(* IEC 61131-3 sources: daoli-st-library/DL_Process (part 44) *)

(* ---- FB_DL_PalletizerLayerSeq.st ---- *)
//==============================================================================
// 功能块：FB_DL_PalletizerLayerSeq ｜ 中文名称：码垛层排布顺控
// 所属子库：DL_Process ｜ 版本：v1.0.1 ｜ 兼容：CODESYS V3.5+ / TwinCAT 3 / 汇川 InoProShop
// 功能描述：码垛机层排布顺控：层容量自算（正交与旋转两取向各算一遍，逐层按本层取向校验）→ 层内位置
//           序列 → 取放指令与夹手完成反馈握手（超时重试一次）→ 层满/垛满判定。
//           奇偶层旋转时偶数层整体旋转 90 度，层内落点由 FC_DL_Affine2Apply 施加旋转
//           矩阵得到（库内低层复用，禁止在本件重写点变换与矩阵乘）。旋转矩阵的元素以
//           VAR CONSTANT 标量常量声明（恒等 1/0、90 度 0/-1/+1），每拍装配成生效阵；
//           平移列恒为 0，运行时平移量（托盘长度）在阵外补偿——阵中不含运行时量，才配
//           得上常量语义（二维数组行主序字面量初始化在三平台可移植性差，故用标量常量
//           装配，避免方言差异）。本件只出位姿与指令，不做轨迹规划、不控夹手电磁阀
//           （执行器归设备层）。
// 开源溯源 (Origin)：道莅原创实现（参考 公开工程惯例 分类与参数域）
// 单位表：托盘与箱体尺寸[mm] / 层高[mm] / 坐标[mm] / 旋转角[度] / 层数与位置序号[个] /
//         取放超时[s] / 扫描间隔[ms] / 垛计数[垛]
// 错误码表：16#0005_0408 信息级（末层不满垛，留空位，不置 bError）/ 16#0005_0409 信息级
//           （取放超时首次重试，不置 bError）/ 16#0005_034E 故障级（层容量不足或箱体/
//           托盘尺寸规格不匹配，含尺寸非有限——非有限尺寸即规格不可信，映射见本行）/
//           16#0005_034F 故障级（取放超时重试耗尽，垛型中断，置 bError + 撤指令）/
//           16#0005_0350 故障级兜底（状态机落 ELSE 非法状态，置 bError）。034E 非有限
//           映射的反证句：尺寸非有限与容量不足在现有输出组合下不可观测出差异（均为
//           bError + bPlaceCmd 撤 + bValid 撤 + eState 进 eFault），§3 未给本件独立非有限
//           槽，故显式复用不越段。
// 状态机：E_DL_PalletLayerState（eIdle=0 待机 / eWaitCase=10 等来料 / ePlace=20 出取放
//           指令 / eWaitGrip=30 等夹手反馈 / eLayerEnd=40 层边界 / ePalletEnd=50 垛边界 /
//           eFault=99 故障兜底），CASE 含 ELSE 兜底，ELSE 置 0350 且撤指令、许可撤。
// 边界行为：① 层容量自算：正交取向 floor(托盘长/箱长) x floor(托盘宽/箱宽)、旋转取向
//           floor(托盘长/箱宽) x floor(托盘宽/箱长)，两取向各自校验——nCasePerLayer 超
//           正交容量 → 故障 034E；启用奇偶层旋转时还须不超旋转容量，否则同样 034E
//           （取大者会让旋转层"蒙混过关"，故逐取向验，绝不硬塞）；② 取放超时先重试
//           一次（信息 0409），二次超时 → 故障 034F 并中断垛型；③ 层高累计 Z =
//           (层号 − 1) x 层高，LREAL 承载防溢出；④ 末层不满 → 信息 0408；⑤ bStop 只在
//           层边界与等来料相生效（不在抓取中停，安全侧）；⑥ 失能/停止 → 撤指令 +
//           bValid := FALSE（R72）；⑦ 旋转落点必须走 FC_DL_Affine2Apply（常量纯旋转阵，
//           平移在阵外补偿），点变换件返回不可用 → 034E 并撤指令。
// 修订历史：v1.0.0 2026-11-17 首版（R25 派单 · §4.16，依赖 §4.2 件 FC_DL_Affine2Apply 语义）
//           v1.0.1 2026-11-17 终审修正两处（对外引脚契约零变更）：①旋转层阵外平移量由 fPalletLengthMm
//           改为 (nRowsEff − 1) x fCaseWidthMm（原式整体多推一个箱宽，首行落点越出托盘边界）；
//           ②bPalletDone 取消本相同拍自撤，撤销点移交 eIdle 相（原实现同拍置位又撤位，脉冲永不外显）。
//           层容量口径经总监独立验算：1200x1000 托盘配 400x300 箱体 → 正交 3x3=9、旋转 4x2=8，
//           派单书 §4.16 验收向量①所写「容量 6」为派单算术笔误，本件实现（9）为准。
//==============================================================================
(*------------------------------------------------------------------------------
 * 枚举: E_DL_PalletLayerState（归属 DL_Process，与 FB_DL_PalletizerLayerSeq 同文件）
 *----------------------------------------------------------------------------*)
TYPE E_DL_PalletLayerState :
(
    eIdle      := 0,   // 待机：指令撤，等 bStart / Idle, command dropped, waiting for start
    eWaitCase  := 10,  // 等来料：本层下一格位已算好，等 bCaseReady / Waiting for the next case
    ePlace     := 20,  // 出指令：bPlaceCmd 置位，等夹手动作 / Command issued, gripper acting
    eWaitGrip  := 30,  // 等反馈：等 bGripDone 或超时 / Waiting for feedback or timeout
    eLayerEnd  := 40,  // 层边界：本层放满，允许在此停止 / Layer boundary, a safe stop point
    ePalletEnd := 50,  // 垛边界：整垛完成，垛计数 +1 / Pallet boundary, pallet counter increments
    eFault     := 99   // 故障兜底：规格不匹配/超时耗尽/非法状态 / Fault fallback
);
END_TYPE

(*==============================================================================
 * 功能块: FB_DL_PalletizerLayerSeq
 * 调用约定: 每个扫描周期无条件调用一次；uDeltaTimeMs 必须注入真实任务间隔。
 *============================================================================*)
FUNCTION_BLOCK FB_DL_PalletizerLayerSeq
VAR_INPUT
    nCasePerLayer    : INT;                        // 每层箱数 [个]，须 <= 层容量 / Cases per layer [pcs], must not exceed the capacity
    nLayersPerPallet : INT;                        // 每垛层数 [层]，合法域 1~20 / Layers per pallet [layers], domain 1..20
    fPalletLengthMm  : LREAL;                      // 托盘长度 [mm]，须 > 0 / Pallet length [mm], must be > 0
    fPalletWidthMm   : LREAL;                      // 托盘宽度 [mm]，须 > 0 / Pallet width [mm], must be > 0
    fCaseLengthMm    : LREAL;                      // 箱体长度 [mm]，须 > 0 / Case length [mm], must be > 0
    fCaseWidthMm     : LREAL;                      // 箱体宽度 [mm]，须 > 0 / Case width [mm], must be > 0
    fLayerHeightMm   : LREAL;                      // 层高 [mm]，须 > 0 / Layer height [mm], must be > 0
    bOddLayerRotate  : BOOL;                       // 奇偶层旋转使能（偶数层旋转 90 度）/ Odd/even layer rotation, even layers rotate 90 degrees
    bCaseReady       : BOOL;                       // 来料在位 / Case available at the pick point
    bGripDone        : BOOL;                       // 夹手完成反馈 / Gripper completion feedback
    tGripTimeout     : TIME := T#8S;               // 取放超时 [ms] / Pick-and-place timeout [ms]
    bStart           : BOOL;                       // 启动（取上升沿）/ Start, rising edge
    bStop            : BOOL;                       // 停止（只在层边界与等来料相生效）/ Stop, honoured only at layer boundaries and while waiting
    bReset           : BOOL;                       // 复位，上升沿回待机并清垛计数锁存位 / Reset, rising edge returns to idle
    uDeltaTimeMs     : UDINT;                      // 扫描间隔 [ms]，调用方注入，禁系统时间函数 / Scan interval [ms], caller-injected
END_VAR
VAR_OUTPUT
    nLayerIndex      : INT;                        // 当前层号 [层]，从 1 起 / Current layer index, 1-based
    nPosIndex        : INT;                        // 层内位置序号 [个]，从 1 起 / In-layer position index, 1-based
    fTargetXMm       : LREAL;                      // 目标位 X [mm] / Target X [mm]
    fTargetYMm       : LREAL;                      // 目标位 Y [mm] / Target Y [mm]
    fTargetZMm       : LREAL;                      // 目标位 Z [mm] / Target Z [mm]
    fTargetRotDeg    : LREAL;                      // 目标旋转角 [度]，0 或 90 / Target rotation [deg], 0 or 90
    bPlaceCmd        : BOOL;                       // 取放指令（层放满/故障/停止即撤）/ Pick-and-place command
    bLayerDone       : BOOL;                       // 本层已放满 / Layer completed
    bPalletDone      : BOOL;                       // 整垛完成 / Pallet completed
    nCaseCount       : INT;                        // 本垛已放件数 [件] / Cases placed on this pallet [pcs]
    uPalletCount     : UDINT;                      // 完成垛数 [垛]，饱和 / Completed pallets [pallets], saturating
    eErr             : UDINT;                      // 错误码，0 = 无错，码位 16#0005_0408 起信息级、16#0005_034E 起故障级（分带见错误码表） / Error code, 0 = no error, band info/fault per the code table
    bError           : BOOL;                       // 故障级标志，仅故障级错误置位 / Fault-class flag, set only on fault-level codes
    bValid           : BOOL;                       // 位姿输出可用标志，失能/故障闸显式 FALSE / Pose usable flag, explicit FALSE on disable/fault gates
    eState           : E_DL_PalletLayerState;      // 主状态机当前状态 / Current state of the main state machine
END_VAR
VAR
    fbReset          : R_TRIG;                     // 复位上升沿检测实例 / Reset rising edge detector
    fbStart          : R_TRIG;                     // 启动上升沿检测实例 / Start rising edge detector
    fbTonGrip        : TON;                        // 取放超时定时器实例 / Pick-and-place timeout timer
    afRotZero        : ARRAY[0..2, 0..2] OF LREAL; // 本拍生效旋转矩阵（恒等或 90 度）/ Effective rotation matrix of this scan
    nCapOrtho        : INT;                        // 正交取向层容量 [件] / Capacity with the orthogonal orientation [pcs]
    nCapRot          : INT;                        // 旋转取向层容量 [件] / Capacity with the rotated orientation [pcs]
    nCapEff          : INT;                        // 本层取向容量 [件] / Capacity of the current orientation [pcs]
    nColsEff         : INT;                        // 本层列数 [个] / Columns of this layer [pcs]
    nRowsEff         : INT;                        // 本层行数 [个] / Rows of this layer [pcs]
    nIdx0            : INT;                        // 层内零基位置序号 [—] / Zero-based in-layer index
    nCol             : INT;                        // 本格位列号（1 基）[列] / Column of this cell, 1-based
    nRow             : INT;                        // 本格位行号（1 基）[行] / Row of this cell, 1-based
    nRetryCnt        : INT;                        // 本格位超时重试次数 [次] / Timeout retry count of this cell
    nLoop            : INT;                        // 赋值循环索引 [—] / Assignment loop index
    fLocalXMm        : LREAL;                      // 箱体自身坐标系 X [mm] / X in the case-local frame [mm]
    fLocalYMm        : LREAL;                      // 箱体自身坐标系 Y [mm] / Y in the case-local frame [mm]
    fOutXMm          : LREAL;                      // 点变换结果 X [mm] / Transformed X [mm]
    fOutYMm          : LREAL;                      // 点变换结果 Y [mm] / Transformed Y [mm]
    uApplyErr        : UDINT;                      // 点变换件错误码暂存 / Point-transform error code staging
    bApplyFault      : BOOL;                       // 点变换件故障标志暂存 / Point-transform fault flag staging
    bApplyValid      : BOOL;                       // 点变换件可用标志暂存 / Point-transform usable flag staging
    bApplyOk         : BOOL;                       // 点变换件返回值暂存 / Point-transform return staging
    bLayerRotated    : BOOL;                       // 本层旋转标志 / This layer is rotated
    bSpaceWarn       : BOOL;                       // 末层不满提示标志 / Under-filled top layer hint
    bGripTimedOut    : BOOL;                       // 取放超时命中 / Pick-and-place timeout hit
    bRearm           : BOOL;                       // 定时器重装脉冲（本拍强制 IN 为 FALSE 一拍）/ Timer re-arm pulse, forces IN FALSE for one scan
    bNonFin          : BOOL;                       // 非有限判定中间标志 / Non-finite detection intermediate flag
    bFirstScan       : BOOL := TRUE;               // 上电首拍标志 / First-scan flag
END_VAR
VAR CONSTANT
    DL_PLS_CODE_INFO_1 : UDINT := 16#0005_0408;    // 信息级槽 1（末层不满垛留空位） / info slot 1
    DL_PLS_CODE_INFO_2 : UDINT := 16#0005_0409;    // 信息级槽 2（取放超时重试） / info slot 2
    DL_PLS_CODE_FLT_1  : UDINT := 16#0005_034E;    // 故障级槽 1（容量不足/规格不匹配） / fault slot 1
    DL_PLS_CODE_FLT_2  : UDINT := 16#0005_034F;    // 故障级槽 2（超时重试耗尽） / fault slot 2
    DL_PLS_CODE_FLT_3  : UDINT := 16#0005_0350;    // 故障级槽 3（非法状态兜底） / fault slot 3, illegal-state fallback
    DL_PLS_ROT90       : LREAL := 90.0;            // 旋转层目标角 [度] / Rotated layer angle [deg]
    DL_PLS_LAYER_MIN   : INT := 1;                 // 层数下限 [层] / Layer count floor
    DL_PLS_LAYER_MAX   : INT := 20;                // 层数上限 [层] / Layer count ceiling
    DL_PLS_CELL_MIN    : INT := 1;                 // 层容量下限 [件] / Layer capacity floor [pcs]
    DL_PLS_CNT_MAX     : UDINT := 16#FFFF_FFFE;    // 垛计数饱和值 [垛] / Pallet counter saturation
    DL_PLS_RETRY_MAX   : INT := 1;                 // 超时重试次数上限 [次] / Retry ceiling [times]
    DL_PLS_ZERO        : LREAL := 0.0;             // 零值常量，避免裸字面量 [—] / Zero constant, avoids a bare literal
    DL_PLS_ONE         : LREAL := 1.0;             // 单位常量，齐次项 [—] / Unity constant, homogeneous entry
    DL_PLS_TOL         : LREAL := 1.0E-6;          // 浮点比较容差 [—] / Float comparison tolerance
    DL_PLS_INF         : LREAL := 1.7976931348623157E308; // LREAL 幅值上限，Inf 判据 / LREAL magnitude ceiling
    // 纯旋转常量阵（行主序平铺展开）：恒等映射 / pure rotation constants, row-major flat
    DL_PLS_M_ID_X      : LREAL := 1.0;             // 恒等阵 (0,0) / identity (0,0)
    DL_PLS_M_ID_Y      : LREAL := 1.0;             // 恒等阵 (1,1) / identity (1,1)
    DL_PLS_M_R90_C     : LREAL := -1.0;            // 90 度阵 (0,1) = -1 / rot90 (0,1) = -1
    DL_PLS_M_R90_S     : LREAL := 1.0;             // 90 度阵 (1,0) = +1 / rot90 (1,0) = +1
END_VAR

(*------------------------------------------------------------------------------
 * 段 1｜无条件刷新区（红线 5）：复位/启动沿与超时定时器在任意分支之外周期调用；
 *       定时器 IN 取上拍状态（单拍滞后对 8 s 窗无影响），保证各分支计时链不断流
 *----------------------------------------------------------------------------*)
fbReset(CLK := bReset);                            // 复位沿检测无条件刷新 / reset edge refreshed unconditionally
fbStart(CLK := bStart);                            // 启动沿检测无条件刷新 / start edge refreshed unconditionally
fbTonGrip(IN := (eState = E_DL_PalletLayerState.eWaitGrip) AND (NOT bGripDone)
                AND (NOT bRearm),                  // 重装拍强制 IN 为 FALSE 使定时器复位 / the re-arm scan forces IN FALSE, resetting the timer
          PT := tGripTimeout);                     // 取放超时 [ms] / pick-and-place timeout
IF bRearm THEN
    bRearm := FALSE;                               // 重装脉冲单拍自清（下一拍起重新计时）/ re-arm pulse self-cleared, timing restarts next scan
END_IF

(*------------------------------------------------------------------------------
 * 段 2｜复位沿处理（改写置于沿后，防吞沿 R39）
 *----------------------------------------------------------------------------*)
IF fbReset.Q THEN
    eState := E_DL_PalletLayerState.eIdle;
    eErr   := 16#0000_0000;                        // 复位清码 / reset clears the code
    bError := FALSE;                               // 复位清故障 / reset clears the fault
    nLayerIndex := 0;                              // 层号清 / layer index cleared
    nPosIndex := 0;                                // 位置序号清 / position index cleared
    nCaseCount := 0;                               // 本垛件数清 / pallet case count cleared
    nRetryCnt := 0;                                // 重试计数清 / retry count cleared
    bPlaceCmd := FALSE;                            // 指令撤 / command dropped
    bFirstScan := TRUE;                            // 重新首拍化 / re-initialize first scan
END_IF

(*------------------------------------------------------------------------------
 * 段 3｜非有限输入闸（尺寸类，R79）：映射入 034E（规格不可信，见错误码表反证句）
 *----------------------------------------------------------------------------*)
bNonFin := (fPalletLengthMm <> fPalletLengthMm) OR (ABS(fPalletLengthMm) >= DL_PLS_INF)
        OR (fPalletWidthMm <> fPalletWidthMm) OR (ABS(fPalletWidthMm) >= DL_PLS_INF)
        OR (fCaseLengthMm <> fCaseLengthMm) OR (ABS(fCaseLengthMm) >= DL_PLS_INF)
        OR (fCaseWidthMm <> fCaseWidthMm) OR (ABS(fCaseWidthMm) >= DL_PLS_INF)
        OR (fLayerHeightMm <> fLayerHeightMm) OR (ABS(fLayerHeightMm) >= DL_PLS_INF);   // 尺寸非有限汇总 / dimensions non-finite
IF bNonFin THEN
    eState := E_DL_PalletLayerState.eFault;        // 进故障相 / enter fault state
    eErr   := DL_PLS_CODE_FLT_1;                   // 故障级：规格不可信 / fault: specification untrustworthy
    bError := TRUE;                                // 故障级必置 bError（R45 配对）/ fault-class pairs with bError
    bPlaceCmd := FALSE;                            // 指令撤安全侧 / command dropped, safe side
    bValid := FALSE;                               // 位姿不可用 / poses unusable
    RETURN;
END_IF

(*------------------------------------------------------------------------------
 * 段 4｜尺寸与层数域闸：尺寸非正会致除零与负坐标倒排（先判后除）
 *----------------------------------------------------------------------------*)
IF (fPalletLengthMm <= DL_PLS_TOL) OR (fPalletWidthMm <= DL_PLS_TOL)
   OR (fCaseLengthMm <= DL_PLS_TOL) OR (fCaseWidthMm <= DL_PLS_TOL)
   OR (fLayerHeightMm <= DL_PLS_TOL)
   OR (nLayersPerPallet < DL_PLS_LAYER_MIN) OR (nLayersPerPallet > DL_PLS_LAYER_MAX) THEN
    eState := E_DL_PalletLayerState.eFault;        // 进故障相 / enter fault state
    eErr   := DL_PLS_CODE_FLT_1;                   // 故障级：尺寸/层数域非法 / fault: dimension or layer domain invalid
    bError := TRUE;                                // 故障级必置 bError（R45 配对）/ fault-class pairs with bError
    bPlaceCmd := FALSE;                            // 指令撤安全侧 / command dropped, safe side
    bValid := FALSE;                               // 位姿不可用 / poses unusable
    RETURN;
END_IF

(*------------------------------------------------------------------------------
 * 段 5｜层容量自算（正交与旋转两取向各算一遍）与数量校验：
 *       容量不足绝不硬塞——基本取向与旋转取向都要单独验，取大者不能让旋转层蒙混过关
 *----------------------------------------------------------------------------*)
nCapOrtho := LREAL_TO_INT(fPalletLengthMm / fCaseLengthMm) * LREAL_TO_INT(fPalletWidthMm / fCaseWidthMm);   // 正交取向容量 [件] / orthogonal capacity [pcs]
nCapRot := LREAL_TO_INT(fPalletLengthMm / fCaseWidthMm) * LREAL_TO_INT(fPalletWidthMm / fCaseLengthMm);     // 旋转取向容量 [件] / rotated capacity [pcs]
IF (nCapOrtho < DL_PLS_CELL_MIN) OR (nCapRot < DL_PLS_CELL_MIN) THEN
    eState := E_DL_PalletLayerState.eFault;        // 进故障相 / enter fault state
    eErr   := DL_PLS_CODE_FLT_1;                   // 故障级：任一取向放不下一个箱 / fault: a case does not fit in one orientation
    bError := TRUE;                                // 故障级必置 bError（R45 配对）/ fault-class pairs with bError
    bPlaceCmd := FALSE;                            // 指令撤安全侧 / command dropped, safe side
    bValid := FALSE;                               // 位姿不可用 / poses unusable
    RETURN;
END_IF
IF (nCasePerLayer < DL_PLS_CELL_MIN) OR (nCasePerLayer > nCapOrtho) THEN
    eState := E_DL_PalletLayerState.eFault;        // 进故障相 / enter fault state
    eErr   := DL_PLS_CODE_FLT_1;                   // 故障级：层容量不足/规格不匹配 / fault: layer capacity or specification mismatch
    bError := TRUE;                                // 故障级必置 bError（R45 配对）/ fault-class pairs with bError
    bPlaceCmd := FALSE;                            // 指令撤安全侧 / command dropped, safe side
    bValid := FALSE;                               // 位姿不可用 / poses unusable
    RETURN;
END_IF
IF bOddLayerRotate AND (nCasePerLayer > nCapRot) THEN
    eState := E_DL_PalletLayerState.eFault;        // 进故障相 / enter fault state
    eErr   := DL_PLS_CODE_FLT_1;                   // 故障级：旋转层容量不足（奇偶层旋转必用旋转取向）/ fault: rotated layers cannot hold the count
    bError := TRUE;                                // 故障级必置 bError（R45 配对）/ fault-class pairs with bError
    bPlaceCmd := FALSE;                            // 指令撤安全侧 / command dropped, safe side
    bValid := FALSE;                               // 位姿不可用 / poses unusable
    RETURN;
END_IF

(*------------------------------------------------------------------------------
 * 段 6｜本层取向与列行数：旋转层箱体足迹长宽互换（足迹互换由矩阵变换真实体现）
 *----------------------------------------------------------------------------*)
bLayerRotated := bOddLayerRotate AND (((nLayerIndex MOD 2) = 0) AND (nLayerIndex >= 1));   // 偶数层旋转（层号 1 基）/ even layers rotate
IF bLayerRotated THEN
    fTargetRotDeg := DL_PLS_ROT90;                 // 目标旋转角 90 度 [度] / target rotation 90 degrees
    nColsEff := LREAL_TO_INT(fPalletWidthMm / fCaseLengthMm);    // 旋转层：列沿托盘宽方向 / rotated: columns run along the pallet width
    nRowsEff := LREAL_TO_INT(fPalletLengthMm / fCaseWidthMm);    // 旋转层：行沿托盘长方向 / rotated: rows run along the pallet length
    nCapEff := nCapRot;                            // 本层容量取旋转取向 [件] / capacity of the rotated orientation [pcs]
    afRotZero[0, 0] := DL_PLS_ZERO;                // rot90 (0,0) = 0 / rot90 (0,0) = 0
    afRotZero[0, 1] := DL_PLS_M_R90_C;             // rot90 (0,1) = -1 / rot90 (0,1) = -1
    afRotZero[0, 2] := DL_PLS_ZERO;                // rot90 平移列 x = 0（运行时平移在阵外补偿）/ rot90 translation x = 0, compensated outside
    afRotZero[1, 0] := DL_PLS_M_R90_S;             // rot90 (1,0) = +1 / rot90 (1,0) = +1
    afRotZero[1, 1] := DL_PLS_ZERO;                // rot90 (1,1) = 0 / rot90 (1,1) = 0
    afRotZero[1, 2] := DL_PLS_ZERO;                // rot90 平移列 y = 0 / rot90 translation y = 0
ELSE
    fTargetRotDeg := DL_PLS_ZERO;                  // 正交层不旋转 [度] / orthogonal layer, no rotation
    nColsEff := LREAL_TO_INT(fPalletLengthMm / fCaseLengthMm);   // 正交层：列沿托盘长方向 / orthogonal: columns along the pallet length
    nRowsEff := LREAL_TO_INT(fPalletWidthMm / fCaseWidthMm);     // 正交层：行沿托盘宽方向 / orthogonal: rows along the pallet width
    nCapEff := nCapOrtho;                          // 本层容量取正交取向 [件] / capacity of the orthogonal orientation [pcs]
    afRotZero[0, 0] := DL_PLS_M_ID_X;              // 恒等阵 (0,0) / identity (0,0)
    afRotZero[0, 1] := DL_PLS_ZERO;                // 恒等阵 (0,1) / identity (0,1)
    afRotZero[0, 2] := DL_PLS_ZERO;                // 恒等阵平移 x = 0 / identity translation x = 0
    afRotZero[1, 0] := DL_PLS_ZERO;                // 恒等阵 (1,0) / identity (1,0)
    afRotZero[1, 1] := DL_PLS_M_ID_Y;              // 恒等阵 (1,1) / identity (1,1)
    afRotZero[1, 2] := DL_PLS_ZERO;                // 恒等阵平移 y = 0 / identity translation y = 0
END_IF
FOR nLoop := 0 TO 2 DO
    afRotZero[2, nLoop] := DL_PLS_ZERO;            // 第三行清零 / third row cleared
END_FOR
afRotZero[2, 2] := DL_PLS_ONE;                     // 齐次项 1（仿射语义要求第三行 0/0/1）/ homogeneous entry 1

(*------------------------------------------------------------------------------
 * 段 7｜层内格位解码与旋转落点：点变换走 FC_DL_Affine2Apply（每拍恰好一次，
 *       禁止复制低层矩阵乘）；旋转层再按托盘长度做阵外平移补偿
 *----------------------------------------------------------------------------*)
nIdx0 := nPosIndex - 1;                            // 零基位置序号 / zero-based index
IF nIdx0 < 0 THEN
    nIdx0 := 0;                                    // 负序号防护 / negative-index guard
END_IF
IF nColsEff < DL_PLS_LAYER_MIN THEN
    nColsEff := DL_PLS_LAYER_MIN;                  // 列数下限防护（防除零）/ column floor guard
END_IF
nRow := (nIdx0 / nColsEff) + 1;                    // 行号（1 基）[行] / row number, 1-based
nCol := nIdx0 - ((nRow - 1) * nColsEff) + 1;       // 列号（1 基）[列] / column number, 1-based
fLocalXMm := INT_TO_LREAL(nCol - 1) * fCaseLengthMm;   // 箱体自身坐标 X [mm] / case-local X [mm]
fLocalYMm := INT_TO_LREAL(nRow - 1) * fCaseWidthMm;    // 箱体自身坐标 Y [mm] / case-local Y [mm]
bApplyOk := FC_DL_Affine2Apply(afM := afRotZero,   // 本拍旋转矩阵 [无量纲+mm] / rotation matrix of this scan
                               fX := fLocalXMm,    // 源点 X [mm] / source X [mm]
                               fY := fLocalYMm,    // 源点 Y [mm] / source Y [mm]
                               fOutX => fOutXMm,   // 变换后 X [mm] / transformed X [mm]
                               fOutY => fOutYMm,   // 变换后 Y [mm] / transformed Y [mm]
                               eErr => uApplyErr,  // 下游错误码暂存 / downstream error code staging
                               bError => bApplyFault,   // 下游故障标志暂存 / downstream fault flag staging
                               bValid => bApplyValid);  // 下游可用标志暂存 / downstream usable flag staging
IF (NOT bApplyValid) OR (NOT bApplyOk) THEN
    eState := E_DL_PalletLayerState.eFault;        // 点变换不可用进故障相 / transform unusable enters fault
    eErr   := DL_PLS_CODE_FLT_1;                   // 故障级：落点不可信（归规格不匹配槽，反证句见头注释）/ fault: pose untrustworthy
    bError := TRUE;                                // 故障级必置 bError（R45 配对）/ fault-class pairs with bError
    bPlaceCmd := FALSE;                            // 指令撤安全侧 / command dropped, safe side
    bValid := FALSE;                               // 位姿不可用 / poses unusable
    RETURN;
END_IF
IF bLayerRotated THEN
    // 旋转 90 度后箱体沿托盘长方向的足迹 = 箱宽 fCaseWidthMm。源点旋转得 X' ∈ [-(nRowsEff−1)x箱宽, 0]，
    // 平移量必须取「满排跨度 − 一个足迹」= (nRowsEff − 1) x 箱宽，落点才严格落在 [0, 托盘长 − 箱宽]。
    // v1.0.1 修正：原式加 fPalletLengthMm 会整体多推一个箱宽，首行落点越出托盘边界（1200x1000 / 箱 400x300 时
    // 得 {300,600,900,1200}，最大角 1500 > 1200）；末角对齐后才与正交取向的 0 基足迹约定一致。
    fTargetXMm := fOutXMm + INT_TO_LREAL(nRowsEff - 1) * fCaseWidthMm;   // 旋转层阵外平移补偿（跨度减一个足迹）[mm] / rotated translation, span minus one footprint
    fTargetYMm := fOutYMm;                         // 旋转层 Y 直接取变换值 [mm] / rotated Y as transformed
ELSE
    fTargetXMm := fOutXMm;                         // 正交层 X 直接取变换值 [mm] / orthogonal X as transformed
    fTargetYMm := fOutYMm;                         // 正交层 Y 直接取变换值 [mm] / orthogonal Y as transformed
END_IF
fTargetZMm := INT_TO_LREAL(nLayerIndex - 1) * fLayerHeightMm;   // 层高累计（LREAL 承载）[mm] / layer height accumulation
bSpaceWarn := (nCasePerLayer < nCapEff);            // 本层留空位（末层不满常见）/ empty slots in this layer

(*------------------------------------------------------------------------------
 * 段 8｜超时判定（各格位独立计时，指令撤后定时器自然复位，禁相内累计）
 *----------------------------------------------------------------------------*)
bGripTimedOut := (eState = E_DL_PalletLayerState.eWaitGrip) AND fbTonGrip.Q AND (NOT bGripDone);   // 超时命中 / timeout hit
IF bGripTimedOut AND (nRetryCnt < DL_PLS_RETRY_MAX) THEN
    nRetryCnt := nRetryCnt + 1;                    // 首次超时：重试计数 +1 [次] / first timeout, retry once
    bRearm := TRUE;                                // 定时器重装：下一拍强制 IN 为 FALSE 一拍再重新计时 / re-arm the timer with one FALSE sample
    eState := E_DL_PalletLayerState.ePlace;        // 回出指令相重发（定时器随之复位）/ re-issue, the timer re-arms
    eErr := DL_PLS_CODE_INFO_2;                    // 信息级：取放超时重试 / info: timeout retried
    bError := FALSE;                               // 信息级不置 bError（R45/R101）/ info never raises bError
ELSIF bGripTimedOut AND (nRetryCnt >= DL_PLS_RETRY_MAX) THEN
    bPlaceCmd := FALSE;                            // 二次超时撤指令（安全侧）/ second timeout drops the command
    eState := E_DL_PalletLayerState.eFault;        // 进故障相 / enter fault state
    eErr   := DL_PLS_CODE_FLT_2;                   // 故障级：超时重试耗尽，垛型中断 / fault: retries exhausted, pallet pattern broken
    bError := TRUE;                                // 故障级必置 bError（R45 配对）/ fault-class pairs with bError
    bValid := FALSE;                               // 位姿不可用 / poses unusable
    RETURN;
END_IF

(*------------------------------------------------------------------------------
 * 段 9｜状态机：CASE 含 ELSE 兜底（非法状态 → 0350 + 撤指令 + 许可撤）
 *----------------------------------------------------------------------------*)
CASE eState OF

    E_DL_PalletLayerState.eIdle:
        bPlaceCmd := FALSE;                        // 待机指令撤 / command dropped in idle
        bValid := FALSE;                           // 失能闸显式不可用（R72）/ explicit FALSE on the disable gate
        bLayerDone := FALSE;                       // 层完成标志撤 / layer-done flag withdrawn
        bPalletDone := FALSE;                      // 垛完成标志撤 / pallet-done flag withdrawn
        nLayerIndex := 0;                          // 层号清 / layer index cleared
        nPosIndex := 1;                            // 位置序号预置 1，便于首件定位 / position index preset to 1
        nCaseCount := 0;                           // 本垛件数清 / pallet case count cleared
        eErr := 16#0000_0000;                      // 待机无错 / no error in idle
        bError := FALSE;                           // 待机无故障 / no fault in idle
        IF fbStart.Q THEN
            eState := E_DL_PalletLayerState.eWaitCase;   // 启动上升沿进等来料 / start edge enters waiting
            nLayerIndex := 1;                      // 从第 1 层开始 / start from layer 1
            nPosIndex := 1;                        // 从第 1 位开始 / start from position 1
            nRetryCnt := 0;                        // 重试计数清 / retry count cleared
            bFirstScan := FALSE;                   // 首拍标志清除 / first-scan flag cleared
        END_IF

    E_DL_PalletLayerState.eWaitCase:
        bPlaceCmd := FALSE;                        // 等来料不出指令 / no command while waiting
        bValid := TRUE;                            // 位姿已算好可用 / the pose is ready and usable
        bError := FALSE;                           // 等料相无故障 / no fault while waiting
        eErr := 16#0000_0000;                      // 等料相先清码 / clear the code first
        IF NOT bCaseReady THEN
            IF bSpaceWarn THEN
                eErr := DL_PLS_CODE_INFO_1;        // 信息级：本层留空位提示 / info: empty slots in this layer
            END_IF
        ELSE
            eState := E_DL_PalletLayerState.ePlace;   // 来料在位出指令（退出条件一）/ case ready, first exit
            nRetryCnt := 0;                        // 新格位重试计数清 / retry count cleared for the new cell
        END_IF
        IF bStop THEN
            eState := E_DL_PalletLayerState.eIdle; // 停止只在等来料相生效（安全侧：不在抓取中停，退出条件二）/ stop honoured here only
            bValid := FALSE;                       // 停止闸显式不可用 / explicit FALSE on the stop gate
            bPlaceCmd := FALSE;                    // 指令撤 / command dropped
        END_IF

    E_DL_PalletLayerState.ePlace:
        bPlaceCmd := TRUE;                         // 取放指令置位 / pick-and-place command raised
        bValid := TRUE;                            // 位姿可用 / poses usable
        bError := FALSE;                           // 出指令相无故障（超时已由段 8 处置）/ no fault here, timeouts handled earlier
        IF eErr <> DL_PLS_CODE_INFO_2 THEN
            eErr := 16#0000_0000;                  // 保留重试提示一拍，其余清码 / keep the retry hint for one scan
        END_IF
        eState := E_DL_PalletLayerState.eWaitGrip; // 无条件进等反馈相（指令保持）/ always enter the feedback wait

    E_DL_PalletLayerState.eWaitGrip:
        bPlaceCmd := TRUE;                         // 指令保持到反馈 / command held until feedback
        bValid := TRUE;                            // 位姿可用 / poses usable
        bError := FALSE;                           // 等反馈相无故障 / no fault while waiting
        IF bGripDone THEN
            nCaseCount := nCaseCount + 1;          // 本垛已放件数 +1 [件] / pallet case count increments
            nPosIndex := nPosIndex + 1;            // 位置序号推进 / position index advances
            nRetryCnt := 0;                        // 重试计数清 / retry count cleared
            bPlaceCmd := FALSE;                    // 反馈到即撤指令 / command dropped on feedback
            IF nPosIndex > nCasePerLayer THEN
                eState := E_DL_PalletLayerState.eLayerEnd;   // 本层放满进层边界 / layer full, enter the layer boundary
            ELSE
                eState := E_DL_PalletLayerState.eWaitCase;   // 本层未满等下一件 / next case in the same layer
            END_IF
        END_IF

    E_DL_PalletLayerState.eLayerEnd:
        bPlaceCmd := FALSE;                        // 层边界指令撤 / command dropped at the layer boundary
        bLayerDone := TRUE;                        // 层完成标志置位 / layer-done flag raised
        bValid := TRUE;                            // 状态可用 / status usable
        bError := FALSE;                           // 层边界无故障 / no fault at the boundary
        eErr := 16#0000_0000;                      // 层边界先清码 / clear the code first
        IF bSpaceWarn THEN
            eErr := DL_PLS_CODE_INFO_1;            // 信息级：本层留空位 / info: empty slots in this layer
        END_IF
        IF bStop THEN
            eState := E_DL_PalletLayerState.eIdle; // 层边界是合法停止点（退出条件一）/ the layer boundary is a legal stop point
            bLayerDone := FALSE;                   // 层完成标志撤 / layer-done flag withdrawn
            bValid := FALSE;                       // 停止闸显式不可用 / explicit FALSE on the stop gate
        ELSIF nLayerIndex >= nLayersPerPallet THEN
            eState := E_DL_PalletLayerState.ePalletEnd;   // 末层已满进垛边界（退出条件二）/ last layer done, second exit
        ELSE
            nLayerIndex := nLayerIndex + 1;        // 升层 / next layer
            nPosIndex := 1;                        // 位置序号回 1 / position index rewound
            bLayerDone := FALSE;                   // 层完成标志撤（升层即清）/ layer-done cleared on the layer change
            eState := E_DL_PalletLayerState.eWaitCase;   // 回等来料（退出条件三）/ back to waiting
        END_IF

    E_DL_PalletLayerState.ePalletEnd:
        bPlaceCmd := FALSE;                        // 垛边界指令撤 / command dropped at the pallet boundary
        bPalletDone := TRUE;                       // 垛完成标志置位 / pallet-done flag raised
        bValid := TRUE;                            // 状态可用 / status usable
        bError := FALSE;                           // 垛边界无故障 / no fault at the boundary
        eErr := 16#0000_0000;                      // 垛边界无错 / no error at the boundary
        IF uPalletCount < DL_PLS_CNT_MAX THEN
            uPalletCount := uPalletCount + 1;      // 完成垛数饱和自增 [垛] / saturating pallet increment
        END_IF
        nLayerIndex := 0;                          // 层号回 0（等下次启动）/ layer index reset
        nPosIndex := 1;                            // 位置序号回 1 / position index rewound
        nCaseCount := 0;                           // 本垛件数清 / pallet case count cleared
        // v1.0.1 修正：bPalletDone 在本相置位后不得同拍自撤（同拍置位+撤位 = 脉冲永不外显）。
        // 撤销点统一放在 eIdle 相（下一拍），保证调用方能采到恰好一拍的 TRUE。
        eState := E_DL_PalletLayerState.eIdle;     // 回待机（bPalletDone 由 eIdle 相撤销）/ back to idle, withdrawn by the idle state

    E_DL_PalletLayerState.eFault:
        bPlaceCmd := FALSE;                        // 故障闸撤指令（R72）/ command dropped on the fault gate
        bValid := FALSE;                           // 故障闸显式不可用 / explicit FALSE on the fault gate
        bError := TRUE;                            // 故障级必置 bError（R45 配对）/ fault-class pairs with bError
        bLayerDone := FALSE;                       // 层完成标志撤 / layer-done flag withdrawn
        IF eErr = 16#0000_0000 THEN
            eErr := DL_PLS_CODE_FLT_3;             // 入口无码时按非法状态兜底（R45：bError 必须有对应码）/ illegal-state fallback
        END_IF
        IF bReset THEN
            eState := E_DL_PalletLayerState.eIdle; // 仅复位可退出故障相 / only reset leaves the fault state
        END_IF

    ELSE
        eState := E_DL_PalletLayerState.eFault;    // 非法状态兜底 / illegal-state fallback
        eErr := DL_PLS_CODE_FLT_3;                 // 故障级兜底：非法状态 / fault fallback: illegal state
        bError := TRUE;                            // 故障级必置 bError（R45 配对）/ fault-class pairs with bError
        bPlaceCmd := FALSE;                        // 指令撤安全侧 / command dropped, safe side
        bValid := FALSE;                           // 位姿不可用 / poses unusable
        bLayerDone := FALSE;                       // 层完成标志撤 / layer-done flag withdrawn
        bPalletDone := FALSE;                      // 垛完成标志撤 / pallet-done flag withdrawn

END_CASE
END_FUNCTION_BLOCK

(* ---- FB_DL_PalletizerStation.st ---- *)
// =====================================================================
// FB_DL_PalletizerStation.st
// 码垛整跺工站编排（进箱→分层码放→层完成→缠膜→出跺，逐相超时）
// Palletizer station sequencing FB via I_DL_Cylinder contracts
// 码位: 16#0005_044E ~ 16#0005_0452 (本件独占 5 槽)
// 修改记录: R29 初版 (按 DISPATCH_R29 序 16)
// =====================================================================
// 枚举: E_DL_PalletizerState（归属 Ownership：E_DL_PalletizerState 归属本文件
//       FB_DL_PalletizerStation，全库唯一定义，本件只定义不重声明）
//       R74 说明：全库 Grep 确认该枚举此前零定义处（仅本件引用 + DISPATCH_R29
//       规格文），E052 即由此产生；成员集严格取自本文件实际使用的相位取值，
//       编号与 DISPATCH_R29 序 16 规格一致（eFault 取 99 保证排序末位）。
// =====================================================================
TYPE E_DL_PalletizerState :
(
    eIdle      := 0,    // 空闲待启动 / Idle, waiting for start
    eWaitBox   := 1,    // 进箱等待：等 bBoxPresent / Waiting for box presence
    ePlace     := 2,    // 分层码放：夹爪闭合后升降下压 / Placing, lowering with gripper closed
    eLayerDone := 3,    // 层排布完成等待外部层序件回馈 / Layer done, waiting external feedback
    eStretch   := 4,    // 缠膜等待 / Stretch wrapping wait
    eDischarge := 5,    // 出跺等待通道就绪 / Discharge wait for outlet ready
    eDone      := 6,    // 一跺完成（单拍后回进箱等待）/ Pallet done, back to wait next scan
    eFault     := 99    // 故障锁存态 / Fault latched state
);
END_TYPE

// =====================================================================
FUNCTION_BLOCK FB_DL_PalletizerStation
VAR_INPUT
    bEnable       : BOOL  := FALSE;    // 使能 / Enable
    bStart        : BOOL  := FALSE;    // 上升沿启动一跺 / Start on edge
    bReset        : BOOL  := FALSE;    // 复位故障 / Reset
    uLayerCount   : USINT  := 10;      // 每跺层数 1~30 / Layers per pallet
    uBoxPerLayer  : USINT  := 6;       // 每层箱数 1~20 / Boxes per layer
    bBoxPresent   : BOOL  := FALSE;    // 入口有箱 / Box present
    bPlaceDone    : BOOL  := FALSE;    // 单箱落位确认 / Box placed
    bLayerDone    : BOOL  := FALSE;    // 层排布完成（外部层序件回馈）/ Layer done
    bStretchDone  : BOOL  := FALSE;    // 缠膜完成 / Stretch done
    bOutReady     : BOOL  := FALSE;    // 出跺通道就绪 / Discharge ready
    bGripClosed   : BOOL  := FALSE;    // 夹爪已闭合反馈 / Gripper closed
    tStepMax      : TIME  := T#20S;    // 单相超时 T#1S~T#300S / Step timeout [s]
END_VAR
VAR_IN_OUT
    iCylGrip      : I_DL_Cylinder;     // 夹爪气缸契约 / Gripper cylinder
    iCylLift      : I_DL_Cylinder;     // 升降气缸契约 / Lift cylinder
END_VAR
VAR_OUTPUT
    eState        : E_DL_PalletizerState;  // 当前相 / State
    uLayerIdx     : USINT;             // 当前层号 0~30 / Layer index
    uBoxIdx       : USINT;             // 当前层内箱号 0~20 / Box index
    bBusy         : BOOL;              // 运行中 / Busy
    bDone         : BOOL;              // 一跺完成（单拍）/ Pallet done pulse
    eErr          : UDINT;             // 错误码 / Error code
END_VAR
VAR
    rtrigStart    : R_TRIG;            // 启动沿检测（无条件刷新）/ Start edge detector
    tonStep       : TON;               // 本相超时定时器（每相进入时重置，禁跨相复用 R21）/ Step timer, reset per phase entry
    bStepTimerOn  : BOOL;              // 相内定时使能 / Phase timer enable
    bLockoutLatch : BOOL := FALSE;     // 联锁错锁存 / Interlock fault latch
    tStepMaxS     : REAL;              // 超时秒值 / Timeout seconds [s]
    xFirstScan    : BOOL  := TRUE;     // 首扫标记 / First-scan flag
END_VAR

// ---------------------------------------------------------------------
// 代码位表（本件独占，勿复用）:
//   16#0005_044E 信息 帧内正常运行
//   16#0005_044F 故障 tStepMax 非法 / 气缸接口未就绪
//   16#0005_0450 故障 uLayerCount=0 / uBoxPerLayer=0 / bEnable 期 iCylGrip.bError
//   16#0005_0451 信息 单相超时 → 停在当前相、bBusy=FALSE
//   16#0005_0452 故障 ePlace 相内 bGripClosed=FALSE（联锁）或跺中途 bReset → 锁存
// ---------------------------------------------------------------------

// ---- 超时秒值 / Timeout seconds ----
tStepMaxS := TIME_TO_REAL(tStepMax) / 1000.0;   // 秒值 / Seconds [s]

// ---- 启动沿检测（无条件刷新）/ Start edge, unconditional ----
rtrigStart(CLK := bStart);      // 沿检测 / Edge detection

// ---- 超时与接口合法性闸 / Timeout and interface validity gate ----
IF (tStepMax = T#0MS) OR (tStepMaxS < 1.0) OR (tStepMaxS > 300.0)
   OR (iCylGrip = 0) OR (iCylLift = 0) THEN    // 接口引用未注入判定（引用为空判零口径）/ Interface reference not injected, null-reference test
    eState := E_DL_PalletizerState.eFault;  // 故障态 / Fault
    bBusy := FALSE;             // 停止运行 / Not busy
    eErr := 16#0005_044F;       // 故障码 / Fault code
    RETURN;                     // 本拍结束 / End of cycle
END_IF

// ---- 组态错闸（含气缸执行器错）/ Configuration and actuator fault gate ----
IF (uLayerCount = 0) OR (uBoxPerLayer = 0) OR (bEnable AND iCylGrip.bFault) THEN
    eState := E_DL_PalletizerState.eFault;  // 故障态 / Fault
    bBusy := FALSE;             // 停止运行 / Not busy
    eErr := 16#0005_0450;       // 故障码 / Fault code
    RETURN;                     // 本拍结束 / End of cycle
END_IF

// ---- 首扫初始化（R16 首扫纪律）/ First-scan initialization ----
IF xFirstScan THEN
    eState := E_DL_PalletizerState.eIdle;   // 空闲 / Idle
    uLayerIdx := 0;             // 层号清零 / Layer cleared
    uBoxIdx := 0;               // 箱号清零 / Box cleared
    bDone := FALSE;             // 脉冲复位 / Pulse reset
    xFirstScan := FALSE;        // 清标记 / Clear flag
END_IF

// ---- 完成脉冲单拍化 / Done pulse one-cycle ----
IF bDone THEN
    bDone := FALSE;             // 下一拍清 / Clear next cycle
END_IF

// ---- 使能撤销：气缸回安全位（夹爪保持、升降下落）/ Disable: cylinders to safe side ----
IF NOT bEnable THEN
    iCylGrip.CmdStop();         // 夹爪保持（接口语义：CmdStop 双线圈全断保持位置）/ Gripper hold via CmdStop
    iCylLift.CmdRetract();      // 升降下落（接口语义：缩回=下落）/ Lift lower = retract
    eState := E_DL_PalletizerState.eIdle;   // 空闲 / Idle
    uLayerIdx := 0;             // 层号清零 / Layer cleared
    uBoxIdx := 0;               // 箱号清零 / Box cleared
    bBusy := FALSE;             // 停止运行 / Not busy
    bLockoutLatch := FALSE;     // 锁存复位 / Latch reset
    eErr := 16#0005_044E;       // 信息级：空闲 / Info: idle
    bStepTimerOn := FALSE;      // 相定时关 / Timer off
    RETURN;                     // 本拍结束 / End of cycle
END_IF

// ---- 故障锁存路径（联锁错/非法复位）/ Fault latch path ----
IF bLockoutLatch THEN
    eState := E_DL_PalletizerState.eFault;  // 故障态 / Fault
    bBusy := FALSE;             // 停止运行 / Not busy
    eErr := 16#0005_0452;       // 故障码回放 / Fault code replay
    IF bReset THEN
        bLockoutLatch := FALSE;     // 解除锁存 / Release latch
        // 未完成跺强制从进箱等待重起并清层号 / Restart from wait, clear indices
        eState := E_DL_PalletizerState.eWaitBox;    // 回进箱等待 / Back to wait
        uLayerIdx := 0;         // 清层号 / Clear layer
        uBoxIdx := 0;           // 清箱号 / Clear box
    END_IF
    RETURN;                     // 本拍结束 / End of cycle
END_IF

// ---- 跺中途非法复位 → 锁存 / Illegal reset mid-pallet → latch ----
IF bReset AND bBusy THEN
    bLockoutLatch := TRUE;      // 锁存 / Latch
    eState := E_DL_PalletizerState.eFault;  // 故障态 / Fault
    bBusy := FALSE;             // 停止运行 / Not busy
    eErr := 16#0005_0452;       // 故障码 / Fault code
    RETURN;                     // 本拍结束 / End of cycle
END_IF

// ---- 空闲态受理启动沿 / Idle accepts start edge ----
IF (eState = E_DL_PalletizerState.eIdle) OR (eState = E_DL_PalletizerState.eWaitBox) THEN
    eErr := 16#0005_044E;       // 信息级：正常 / Info: normal
    IF rtrigStart.Q AND (eState = E_DL_PalletizerState.eIdle) THEN
        eState := E_DL_PalletizerState.eWaitBox;    // 进入进箱等待 / Go to wait
        uLayerIdx := 1;         // 层号从 1 起 / Layer starts at 1
        uBoxIdx := 1;           // 箱号从 1 起 / Box starts at 1
        bBusy := TRUE;          // 运行 / Busy
        bStepTimerOn := FALSE;  // 相定时未启 / Timer off
    END_IF
END_IF

// ---- 相超时定时器（每相进入时重置，R21 禁跨相复用）/ Step timer, reset per phase entry ----
tonStep(IN := bStepTimerOn, PT := tStepMax);    // 无条件刷新 / Unconditional refresh
IF bStepTimerOn AND tonStep.Q THEN
    bStepTimerOn := FALSE;      // 相定时关 / Timer off
    bBusy := FALSE;             // 停在当前相 / Stay in current phase
    eErr := 16#0005_0451;       // 信息级：单相超时 / Info: step timeout
    RETURN;                     // 不自动跳步 / No auto skip
END_IF

// ---- 状态机 / State machine ----
CASE eState OF

    E_DL_PalletizerState.eIdle: // 空闲态 / Idle
        bBusy := FALSE;         // 非运行 / Not busy
        bStepTimerOn := FALSE;  // 定时关 / Timer off

    E_DL_PalletizerState.eWaitBox:  // 进箱等待 / Wait for box
        bBusy := TRUE;          // 运行 / Busy
        bStepTimerOn := TRUE;   // 相定时启 / Timer on
        IF bBoxPresent THEN
            // 有箱：夹爪闭合准备抓取 / Box present: close gripper
            iCylGrip.CmdExtend();   // 夹爪闭合（接口语义：伸出=夹紧）/ Gripper close = extend
            bStepTimerOn := FALSE;  // 相定时重置 / Timer reset
            eState := E_DL_PalletizerState.ePlace;  // 进入码放相 / Go to place
            tonStep(IN := FALSE, PT := tStepMax);   // 相进入重置（R21）/ Reset on entry
        END_IF

    E_DL_PalletizerState.ePlace:    // 分层码放 / Placing
        bBusy := TRUE;          // 运行 / Busy
        bStepTimerOn := TRUE;   // 相定时启 / Timer on
        // 联锁：夹爪未闭合就允许下压 → 故障锁存 / Interlock: no grip while lowering
        IF NOT bGripClosed THEN
            bLockoutLatch := TRUE;  // 锁存 / Latch
            eErr := 16#0005_0452;   // 故障码 / Fault code
            RETURN;             // 本拍结束 / End of cycle
        END_IF
        iCylLift.CmdRetract();  // 升降下压（接口语义：缩回=下压）/ Lift press = retract
        IF bPlaceDone THEN
            iCylGrip.CmdRetract();   // 夹爪松开（接口语义：缩回=松开）/ Gripper open = retract
            uBoxIdx := uBoxIdx + 1; // 箱号递增 / Box increment
            IF uBoxIdx > uBoxPerLayer THEN
                uBoxIdx := 1;   // 显式回绕到层首 / Wrap to layer first
                bStepTimerOn := FALSE;  // 相定时重置 / Timer reset
                eState := E_DL_PalletizerState.eLayerDone;  // 层完成相 / Layer done phase
                tonStep(IN := FALSE, PT := tStepMax);   // 相进入重置 / Reset on entry
            ELSE
                // 还有箱：回进箱等待取下一箱 / More boxes: back to wait
                bStepTimerOn := FALSE;  // 相定时重置 / Timer reset
                eState := E_DL_PalletizerState.eWaitBox;    // 回等待 / Back to wait
                tonStep(IN := FALSE, PT := tStepMax);   // 相进入重置 / Reset on entry
            END_IF
        END_IF

    E_DL_PalletizerState.eLayerDone:    // 层完成等待 / Layer done wait
        bBusy := TRUE;          // 运行 / Busy
        bStepTimerOn := TRUE;   // 相定时启 / Timer on
        IF bLayerDone THEN
            IF uLayerIdx >= uLayerCount THEN
                // 满跺：进入缠膜 / Full pallet: stretch phase
                bStepTimerOn := FALSE;  // 相定时重置 / Timer reset
                eState := E_DL_PalletizerState.eStretch;    // 缠膜相 / Stretch phase
                tonStep(IN := FALSE, PT := tStepMax);   // 相进入重置 / Reset on entry
            ELSE
                uLayerIdx := uLayerIdx + 1;     // 层号递增 / Layer increment
                uBoxIdx := 1;   // 箱号回层首 / Box to first
                bStepTimerOn := FALSE;  // 相定时重置 / Timer reset
                eState := E_DL_PalletizerState.eWaitBox;    // 回进箱等待 / Back to wait
                tonStep(IN := FALSE, PT := tStepMax);   // 相进入重置 / Reset on entry
            END_IF
        END_IF

    E_DL_PalletizerState.eStretch:  // 缠膜等待 / Stretch wait
        bBusy := TRUE;          // 运行 / Busy
        bStepTimerOn := TRUE;   // 相定时启 / Timer on
        IF bStretchDone THEN
            bStepTimerOn := FALSE;  // 相定时重置 / Timer reset
            eState := E_DL_PalletizerState.eDischarge;  // 出跺相 / Discharge phase
            tonStep(IN := FALSE, PT := tStepMax);   // 相进入重置 / Reset on entry
        END_IF

    E_DL_PalletizerState.eDischarge:    // 出跺等待 / Discharge wait
        bBusy := TRUE;          // 运行 / Busy
        bStepTimerOn := TRUE;   // 相定时启 / Timer on
        IF bOutReady THEN
            bStepTimerOn := FALSE;  // 相定时关 / Timer off
            bDone := TRUE;      // 一跺完成脉冲 / Done pulse
            eState := E_DL_PalletizerState.eDone;   // 完成态 / Done state
            tonStep(IN := FALSE, PT := tStepMax);   // 定时重置 / Reset
        END_IF

    E_DL_PalletizerState.eDone:     // 完成态（下一拍回等待）/ Done, back next cycle
        bBusy := FALSE;         // 非运行 / Not busy
        eState := E_DL_PalletizerState.eWaitBox;    // 回进箱等待 / Back to wait
        uLayerIdx := 0;         // 层号清零 / Layer cleared
        uBoxIdx := 0;           // 箱号清零 / Box cleared

    E_DL_PalletizerState.eFault:    // 故障态 / Fault
        bBusy := FALSE;         // 非运行 / Not busy
        bStepTimerOn := FALSE;  // 定时关 / Timer off

    ELSE                        // 非法状态拦截 / Illegal state interception
        eState := E_DL_PalletizerState.eFault;  // 落故障态 / Fall to fault
        bBusy := FALSE;         // 非运行 / Not busy
        eErr := 16#0005_044E;   // 信息级（状态机兜底非故障源）/ Info
END_CASE

// ---- 气缸执行器错实时登记 / Actuator error live registration ----
IF iCylGrip.bFault OR iCylLift.bFault THEN
    eErr := 16#0005_0450;       // 故障码 / Fault code
    eState := E_DL_PalletizerState.eFault;  // 故障态 / Fault
    bBusy := FALSE;             // 停止运行 / Not busy
END_IF

END_FUNCTION_BLOCK

(* ---- FB_DL_PalletLabelVerify.st ---- *)
(*==============================================================================
 * 组件名称 (Component)  : FB_DL_PalletLabelVerify
 * 所属子库 (Sublibrary) : DL_Process
 * 当前版本 (Version)    : 1.0.0
 * 兼容性 (Platform)     : CODESYS 3.5+ / TwinCAT 3 / 汇川 InoProShop / 施耐德 Machine Expert
 *                         仅依赖 Standard.library（R_TRIG / MID / LEN / MOD），零厂商私有库
 * 功能描述 (Function)   : 托盘标签 EAN-13 校验与错标拦截。触发沿对 13 位码
 *                         串做三段校验：① 长度 = 13；② 逐位数字字符域；
 *                         ③ 校验位复算（位 1..12 权 1/3 交替，chk = (10 -
 *                         Σ mod 10) mod 10 对位 13）。任一段失败即拦截
 *                         bReject 并给出独立错因分码（R190）。与 Crc16Modbus/
 *                         StringTrim（原子件）分工：本件是分段+复算+拦截的
 *                         组合契约件。
 * 来源标签 (Origin)     : ROADMAP §19.4 R12 池（L832），自研 clean-room
 * 边界语义 (Boundary)   : ① 字符提取用标准 MID（下标 1..13 结构性有界）；
 *                         ② 非数字字符在逐位域闸拦截（短路计错即停扫描）；
 *                         ③ 校验复算的 MOD 只作用于非负 INT 和（结构性安全）；
 *                         ④ 长度闸先行：长度不对不进逐位扫描（省时且防越界）。
 * 输出语义 (Fallback)   : 【R191】bEnable = FALSE → 判定输出冻结保持；eFault
 *                         相（非法相位兜底）→ 冻结 + bError = TRUE；校验失败
 *                         是业务结果不是 FB 故障（不置 bError）。
 * 码位     (Codes)      : 按 R297 范式零 16# 码位硬编码；错误出口 BOOL+ENUM(eCause)。
 * 红线自检 (Redline)    : 7 项红线已自检：R1 零全局 ✓｜R2 零物理地址 ✓｜R3 纯 IEC ✓
 *                         R4 越界（MID 有界）/MOD 非负 ✓｜R5 双语同行注释 ✓
 *                         R6 CASE 带 ELSE 兜底迁 eFault ✓｜R7 R_TRIG 段 0 无条件刷新 ✓
 * 验收向量 (Acceptance) : V1 sCode='4006381333931' → 三段全过，bVerifyOk=TRUE
 *                         （EAN-13 公开标准样例码）；
 *                         V2 sCode='4006381333930'（末位错）→ bChkOk=FALSE，
 *                         eErrKind=eChk，bReject 单拍；
 *                         V3 sCode='40063'（长度 5）→ eErrKind=eLen，不进逐位扫描。
 * 修订历史 (Revision)   : 2026-11-20  v1.0.0  R51 首版（批 3 · 序号 11）
 *==============================================================================*)
TYPE E_DL_PlvErrKind :
(
    eOk    := 0,                             (* 校验通过 / Verify pass *)
    eLen   := 1,                             (* 长度不为 13 / Length fault *)
    eChar  := 2,                             (* 存在非数字字符 / Non-digit char *)
    eChk   := 3                              (* 校验位复算不符 / Check-digit mismatch *)
);
END_TYPE

TYPE E_DL_PlvState :
(
    eIdle  := 0,                             (* 待使能 / Idle *)
    eCheck := 10,                            (* 校验运行 / Check run *)
    eFault := 90                             (* 故障锁存相 / Fault latched phase *)
);
END_TYPE

TYPE E_DL_PlvCause :
(
    eNone     := 0,                          (* 无故障成因 / No cause *)
    ePhaseBad := 3                           (* 非法相位兜底 / Illegal phase fallback *)
);
END_TYPE

FUNCTION_BLOCK FB_DL_PalletLabelVerify
VAR_INPUT
    sCode     : STRING := '';                (* 待校验码串（触屏/扫码器接入）[-] / Code string *)
    bVerifyReq: BOOL := FALSE;               (* 校验触发电平（上升沿执行）[-] / Verify trigger *)
    bEnable   : BOOL := TRUE;                (* 使能 [-] / Enable *)
    bReset    : BOOL := FALSE;               (* 复位命令，上升沿清全部 [-] / Reset command *)
END_VAR
VAR_OUTPUT
    bVerifyOk : BOOL;                        (* 三段校验全过（保持到下个触发沿）[-] / Verify verdict *)
    bLenOk    : BOOL;                        (* 长度段结果 [-] / Length verdict *)
    bCharOk   : BOOL;                        (* 字符域段结果 [-] / Char verdict *)
    bChkOk    : BOOL;                        (* 校验位段结果 [-] / Check-digit verdict *)
    eErrKind  : E_DL_PlvErrKind;             (* 错因分码（信息级逐拍重算，R189） / Error kind *)
    bReject   : BOOL;                        (* 拦截单拍位 [-] / Reject pulse *)
    nVerifyCnt: UDINT;                       (* 累计校验次数 [次] / Verify count *)
    eState    : E_DL_PlvState;               (* 状态出口 / State outlet *)
    eCause    : E_DL_PlvCause;               (* 故障成因出口 / Fault cause outlet *)
    bError    : BOOL;                        (* 故障锁存标志 [-] / Fault latch flag *)
END_VAR
VAR
    _eState   : E_DL_PlvState := E_DL_PlvState.eIdle;     (* 内部相位（CASE 唯一写入目标） / Internal phase *)
    _eCause   : E_DL_PlvCause := E_DL_PlvCause.eNone;     (* 故障成因锁存量 / Latched cause *)
    rtReq     : R_TRIG;                      (* 触发沿实例，段 0 无条件调用 / Trigger edge instance *)
    rtReset   : R_TRIG;                      (* 复位沿实例，段 0 无条件调用 / Reset edge instance *)
    _nLen     : INT;                         (* 码串长度工作量 [字符] / Length work *)
    _i        : INT;                         (* 位扫描游标（每趟重置，R227）[-] / Digit cursor *)
    _c        : STRING(1);                   (* 当前位单字符工作量 [-] / Current char work *)
    _nD       : INT;                         (* 当前位数值工作量 [-] / Digit value work *)
    _nSum     : INT;                         (* 加权和工作量 [-] / Weighted sum work *)
    _nChk     : INT;                         (* 复算校验位工作量 [-] / Recomputed check work *)
    _bCharBad : BOOL;                        (* 本串含非数字当拍量 [-] / Non-digit flag *)
    _nVerC    : UDINT;                       (* 校验计数锁存 [次] / Verify count latch *)
    _bFault   : BOOL;                        (* 故障锁存位 / Latched fault bit *)
END_VAR
VAR CONSTANT
    DL_PLV_EANLEN : INT := 13;               (* EAN-13 码长 [字符] / EAN-13 length *)
END_VAR

(* —— 段 0：沿实例无条件刷新（R228A） —— *)
rtReq(CLK := bVerifyReq);                    (* 触发沿每拍必调 / Trigger edge every scan *)
rtReset(CLK := bReset);                      (* 复位沿每拍必调 / Reset edge every scan *)

(* —— 段 1：单拍量预清零（R107） —— *)
bReject := FALSE;                            (* 拦截脉冲预清，唯一分支置位 / Reject preset *)
eErrKind := E_DL_PlvErrKind.eOk;             (* 错因预置通过（判定分支覆盖） / Err kind preset *)

(* —— 段 2：复位沿处理（作用域：清故障 + 清判定出口 + 清计数 + 迁 eIdle，R283 逐项声明） —— *)
IF rtReset.Q THEN
    _bFault := FALSE;                        (* 清故障锁存 / Clear fault *)
    _eCause := E_DL_PlvCause.eNone;          (* 清成因 / Clear cause *)
    bVerifyOk := FALSE;                      (* 清判定出口 / Clear verdict outlet *)
    bLenOk := FALSE;                         (* 清长度段出口 / Clear len outlet *)
    bCharOk := FALSE;                        (* 清字符段出口 / Clear char outlet *)
    bChkOk := FALSE;                         (* 清校验段出口 / Clear chk outlet *)
    _nVerC := 0;                             (* 清计数 / Clear count *)
    _eState := E_DL_PlvState.eIdle;          (* 迁待机相 / Back to idle *)
END_IF

(* —— 段 4：CASE 主状态机（ELSE 兜底迁 eFault，红线 6） —— *)
CASE _eState OF
    E_DL_PlvState.eIdle:                     (* 待机相 / Idle *)
        IF bEnable AND NOT _bFault THEN
            _eState := E_DL_PlvState.eCheck; (* 进入校验 / Enter check *)
        END_IF
    E_DL_PlvState.eCheck:                    (* 校验相：三段串行闸 / Check *)
        IF NOT bEnable THEN
            _eState := E_DL_PlvState.eIdle;  (* 失能回待机 / Back to idle *)
        ELSIF rtReq.Q THEN                   (* 触发沿执行 / On trigger edge *)
            _nVerC := _nVerC + 1;            (* 校验计数（UDINT 回绕工程安全） / Count verify *)
            _nLen := LEN(sCode);             (* 长度段（标准 LEN） / Length stage *)
            bLenOk := (_nLen = DL_PLV_EANLEN);   (* 长度判定 / Length verdict *)
            bCharOk := FALSE;                (* 字符段预置（短路语义：长度错时保持 FALSE） / Char preset *)
            bChkOk := FALSE;                 (* 校验段预置 / Chk preset *)
            bVerifyOk := FALSE;              (* 总判定预置（各通过段刷新） / Verdict preset *)
            IF bLenOk THEN
                _i := 1;                     (* 位游标重置（R227） / Digit cursor reset *)
                _bCharBad := FALSE;          (* 非数字标志重置 / Non-digit reset *)
                _nSum := 0;                  (* 加权和重置 / Sum reset *)
                WHILE _i <= 12 DO            (* 位 1..12：字符域 + 加权和（MID 下标 1..13 有界，边界①） / Digits 1..12 *)
                    _c := MID(sCode, 1, _i); (* 单字符提取（标准 MID） / Extract char *)
                    IF _c = '0' THEN
                        _nD := 0;            (* 数字 0 / Digit 0 *)
                    ELSIF _c = '1' THEN
                        _nD := 1;            (* 数字 1 / Digit 1 *)
                    ELSIF _c = '2' THEN
                        _nD := 2;            (* 数字 2 / Digit 2 *)
                    ELSIF _c = '3' THEN
                        _nD := 3;            (* 数字 3 / Digit 3 *)
                    ELSIF _c = '4' THEN
                        _nD := 4;            (* 数字 4 / Digit 4 *)
                    ELSIF _c = '5' THEN
                        _nD := 5;            (* 数字 5 / Digit 5 *)
                    ELSIF _c = '6' THEN
                        _nD := 6;            (* 数字 6 / Digit 6 *)
                    ELSIF _c = '7' THEN
                        _nD := 7;            (* 数字 7 / Digit 7 *)
                    ELSIF _c = '8' THEN
                        _nD := 8;            (* 数字 8 / Digit 8 *)
                    ELSIF _c = '9' THEN
                        _nD := 9;            (* 数字 9 / Digit 9 *)
                    ELSE
                        _nD := -1;           (* 非数字哨兵 / Non-digit sentinel *)
                        _bCharBad := TRUE;   (* 置非数字标志 / Set flag *)
                    END_IF
                    IF (NOT _bCharBad) AND (_nD >= 0) THEN   (* 域内才累计（短路计错即停，边界②） / Accumulate in-domain *)
                        IF (_i MOD 2) = 1 THEN
                            _nSum := _nSum + _nD;        (* 奇位权 1 / Odd weight 1 *)
                        ELSE
                            _nSum := _nSum + 3 * _nD;    (* 偶位权 3 / Even weight 3 *)
                        END_IF
                    END_IF
                    _i := _i + 1;            (* 游标递进 / Cursor advance *)
                END_WHILE
                bCharOk := NOT _bCharBad;    (* 字符段判定 / Char verdict *)
                IF bCharOk THEN
                    _nChk := (10 - (_nSum MOD 10)) MOD 10;   (* 校验位复算（Σ >= 0 非负，MOD 结构性安全，边界③） / Recompute check digit *)
                    _c := MID(sCode, 1, 13); (* 第 13 位字符 / 13th char *)
                    IF ((_nChk = 0) AND (_c = '0')) OR ((_nChk = 1) AND (_c = '1'))
                       OR ((_nChk = 2) AND (_c = '2')) OR ((_nChk = 3) AND (_c = '3'))
                       OR ((_nChk = 4) AND (_c = '4')) OR ((_nChk = 5) AND (_c = '5'))
                       OR ((_nChk = 6) AND (_c = '6')) OR ((_nChk = 7) AND (_c = '7'))
                       OR ((_nChk = 8) AND (_c = '8')) OR ((_nChk = 9) AND (_c = '9')) THEN
                        bChkOk := TRUE;      (* 校验位匹配 / Chk match *)
                    END_IF
                END_IF
                bVerifyOk := bChkOk;         (* 总判定（长度与字符段已过） / Verdict *)
                IF NOT bLenOk THEN
                    eErrKind := E_DL_PlvErrKind.eLen;    (* 错因：长度 / Kind: length *)
                ELSIF NOT bCharOk THEN
                    eErrKind := E_DL_PlvErrKind.eChar;   (* 错因：字符（独立分码，R190） / Kind: char *)
                ELSIF NOT bChkOk THEN
                    eErrKind := E_DL_PlvErrKind.eChk;    (* 错因：校验位（独立分码） / Kind: chk *)
                END_IF
                bReject := NOT bVerifyOk;    (* 拦截单拍（错标即拦） / Reject on fail *)
            ELSE
                eErrKind := E_DL_PlvErrKind.eLen;    (* 长度闸先行（边界④） / Length gate first *)
                bReject := TRUE;             (* 拦截单拍 / Reject pulse *)
            END_IF
        END_IF
    E_DL_PlvState.eFault:                    (* 故障相：冻结保持，仅复位沿出 / Fault *)
        ;                                    (* 锁存回放（R28） / Replay from latch *)
    ELSE                                     (* 非法相位兜底迁安全态 / Illegal phase fallback *)
        _eState := E_DL_PlvState.eFault;     (* 迁故障相 / To fault *)
        _bFault := TRUE;                     (* 同步锁存 / Latch *)
        _eCause := E_DL_PlvCause.ePhaseBad;  (* 成因：非法相位 / Cause: illegal phase *)
END_CASE

(* —— 段 5：出口映射（bError/eState 同源，R191） —— *)
nVerifyCnt := _nVerC;                        (* 校验计数出口 / Count outlet *)
bError := _bFault;                           (* 故障标志镜像（业务拒绝不置 bError，输出语义声明） / Fault flag mirror *)
eState := _eState;                           (* 状态出口 / State outlet *)
eCause := _eCause;                           (* 成因出口 / Cause outlet *)
END_FUNCTION_BLOCK

(* ---- FB_DL_PalletZoneMerge.st ---- *)
// =====================================================================
// FB_DL_PalletZoneMerge.st
// 码垛前多线合流积放（多区占用去抖 + 释放互斥节流 + 双模式仲裁 + 上区补跑）
// Pallet merge accumulation across zones with mutex release throttling
// 所属子库: DL_Process    版本: v1.0.0    兼容: CODESYS V3.5+ / TwinCAT 3 / 汇川 InoProShop
// 码位: 16#0005_0471 ~ 16#0005_0475 (本件独占 5 槽, 勿复用)
// 溯源: 道莅 clean-room 防御性实现
//       来源组标签: packaging, conveyor, merge, accumulation
// 修改记录: R30 初版 (ROUND_PLAN_R30 序 8)
// 语义声明: 释放输出为单拍脉冲（当拍自清）, 下游合流区须自行锁存接续;
//           上区补跑语义: 被节流/等待的占用区在条件恢复后按同一仲裁律
//           逐拍继续放出, 不丢件; 光电闪断经关断延时去抖, 短闪不丢占用
// =====================================================================
FUNCTION_BLOCK FB_DL_PalletZoneMerge
VAR_INPUT
    bEnable    : BOOL  := FALSE;    // 使能 / Enable
    abZiOcc    : ARRAY[1..4] OF BOOL;   // 各区光电占用信号 / Zone photoeye occupancy
    bMergeReq  : BOOL  := FALSE;    // 合流释放请求 / Merge release request
    tZiGapMin  : TIME  := T#500MS;  // 相邻两次释放最小间隔, 兼作占用去抖保持窗 / Min release gap, also occupancy hold
    uMergeMode : USINT := 1;        // 合流模式: 1 = 顺序, 2 = 先到先走 / Merge mode
END_VAR
VAR_OUTPUT
    abZiRelease : ARRAY[1..4] OF BOOL;  // 各区释放脉冲输出（单拍自清）/ Zone release pulse, one cycle
    bMergeBusy  : BOOL := FALSE;    // 合流进行中（有请求且有占用区等待）/ Merge busy
    uReleaseSeq : USINT := 0;       // 累计释放次数台账 / Cumulative release count
    eErr        : UDINT := 16#0005_0471;  // 错误码 / Error code
END_VAR
VAR
    aTofOcc    : ARRAY[1..4] OF TOF;    // 各区占用关断延时去抖, 每拍无条件刷新 / Zone occupancy TOF debounce, refreshed every cycle
    aRtrOcc    : ARRAY[1..4] OF R_TRIG; // 各区占用到达沿检测, 每拍无条件刷新 / Zone arrival edges, refreshed every cycle
    tonGap     : TON;               // 释放节流窗定时器, 每拍无条件刷新 / Release throttle timer, refreshed every cycle
    abOccDb    : ARRAY[1..4] OF BOOL;   // 去抖后的区占用 / Debounced occupancy
    auiArrSeq  : ARRAY[1..4] OF USINT;  // 各区到达序号, 0 = 未登记 / Zone arrival sequence, 0 = none
    uArrCnt    : USINT := 0;        // 到达序号累计器 / Arrival sequence counter
    bGapHold   : BOOL := FALSE;     // 节流窗保持标志 / Throttle window hold flag
    bModeOk    : BOOL := FALSE;     // 合流模式合法标记 / Merge mode legal flag
    uSel       : USINT := 0;        // 本拍选中释放区号 / Selected zone this cycle
    uMinSeq    : USINT := 0;        // 最小到达序号临时量 / Min arrival sequence temporary
    uZi        : INT   := 1;        // 1..4 数组下标 / Array subscript 1..4
END_VAR

// ---------------------------------------------------------------------
// 代码位表（本件独占, 勿复用）:
//   16#0005_0471 信息 合流正常（空闲或释放完成）
//   16#0005_0472 故障 合流模式非法冻结（模式值非 1 或 2, 冻结全部释放输出）,
//                解除式 = 模式值恢复合法域
//   16#0005_0473 信息 请求悬空（有合流请求但暂无去抖占用区可释放）
//   16#0005_0474 信息 释放节流窗激活（距上次释放不足最小间隔）
//   16#0005_0475 信息 待机未使能
// ---------------------------------------------------------------------

// ---- 模式合法性 / Merge mode legality ----
IF (uMergeMode = 1) OR (uMergeMode = 2) THEN
    bModeOk := TRUE;                // 合法模式 / Legal mode
ELSE
    bModeOk := FALSE;               // 非法模式冻结 / Illegal mode frozen
END_IF

// ---- 未使能待机处理 / Standby when disabled ----
IF NOT bEnable THEN
    FOR uZi := 1 TO 4 DO
        auiArrSeq[uZi] := 0;        // 清到达序号 / Clear arrival sequence
    END_FOR
    uArrCnt  := 0;                  // 清序号累计器 / Clear counter
    bGapHold := FALSE;              // 清节流标志 / Clear throttle flag
END_IF

// ---- 去抖与到达沿实例无条件周期刷新（4 实例逐个全刷新, 不进 IF 分支）
//      Unconditional refresh of all 4 TOF and 4 R_TRIG instances ----
FOR uZi := 1 TO 4 DO
    aTofOcc[uZi](IN := abZiOcc[uZi], PT := tZiGapMin);  // 闪断保持: 短于间隔窗的闪断不丢占用 / Flicker hold
    aRtrOcc[uZi](CLK := abZiOcc[uZi]);                  // 到达沿 / Arrival edge
    abOccDb[uZi] := aTofOcc[uZi].Q;                     // 去抖后占用 / Debounced occupancy
END_FOR

// ---- 到达序号登记（先到先走模式的次序依据）/ Arrival sequence registration ----
FOR uZi := 1 TO 4 DO
    IF aRtrOcc[uZi].Q AND (auiArrSeq[uZi] = 0) THEN
        uArrCnt := uArrCnt + 1;     // 序号推进 / Advance sequence
        auiArrSeq[uZi] := uArrCnt;  // 登记该区到达序号 / Register arrival
    END_IF
    IF NOT abOccDb[uZi] THEN
        auiArrSeq[uZi] := 0;        // 占用消失清序号 / Clear sequence on vacancy
    END_IF
END_FOR
// 序号累计器回绕防护: 临近上界按当前占用区号序重排 / Counter wrap protection: renumber by zone order
IF uArrCnt >= 250 THEN
    uArrCnt := 0;                   // 累计器归零 / Reset counter
    FOR uZi := 1 TO 4 DO
        auiArrSeq[uZi] := 0;        // 全清后重排 / Clear then renumber
    END_FOR
    FOR uZi := 1 TO 4 DO
        IF abOccDb[uZi] THEN
            uArrCnt := uArrCnt + 1;
            auiArrSeq[uZi] := uArrCnt;  // 按区号序重排占用区 / Renumber occupied zones
        END_IF
    END_FOR
END_IF

// ---- 释放节流窗定时器无条件刷新 / Unconditional throttle timer refresh ----
tonGap(IN := bGapHold, PT := tZiGapMin);
IF tonGap.Q THEN
    bGapHold := FALSE;              // 节流窗完成, 允许下一次释放 / Window done, allow next release
END_IF

// ---- 释放仲裁: 同拍至多一区（互斥）; 多区请求取最小区号或最先到达区
//      Release arbitration: at most one zone per cycle, mutex guaranteed ----
uSel := 0;                          // 选中区清零 / Clear selection
IF bEnable AND bModeOk AND bMergeReq AND (NOT bGapHold) THEN
    IF uMergeMode = 1 THEN
        // 顺序模式: 升序取最小区号 / Sequential: lowest zone number
        FOR uZi := 1 TO 4 DO
            IF (uSel = 0) AND abOccDb[uZi] THEN
                uSel := INT_TO_USINT(uZi);  // 选中该区 / Select zone
            END_IF
        END_FOR
    ELSE
        // 先到先走模式: 取最小到达序号 / First-arrived: min arrival sequence
        uMinSeq := 0;               // 0 表示尚未找到候选 / 0 = no candidate yet
        FOR uZi := 1 TO 4 DO
            IF abOccDb[uZi] THEN
                IF (uMinSeq = 0) OR (auiArrSeq[uZi] < uMinSeq) THEN
                    uMinSeq := auiArrSeq[uZi];  // 更新最小序号 / Update min sequence
                    uSel := INT_TO_USINT(uZi);  // 选中该区 / Select zone
                END_IF
            END_IF
        END_FOR
    END_IF
END_IF

// ---- 释放执行（单拍脉冲, 选中区置真一拍后由下拍缺省清零）
//      Release execution: one-cycle pulse on selected zone ----
FOR uZi := 1 TO 4 DO
    abZiRelease[uZi] := FALSE;      // 缺省全断 / Default all off
END_FOR
IF (uSel >= 1) AND (uSel <= 4) THEN
    abZiRelease[uSel] := TRUE;      // 选中区发释放脉冲（下标已越界守卫）/ Selected zone release pulse, index guarded
    bGapHold := TRUE;               // 启动节流窗 / Start throttle window
    uReleaseSeq := uReleaseSeq + 1; // 释放台账推进 / Advance release ledger
    auiArrSeq[uSel] := 0;           // 该区序号清零待再到达 / Clear its sequence
END_IF

// ---- 合流忙输出 / Merge busy output ----
bMergeBusy := FALSE;                // 缺省不忙 / Default idle
FOR uZi := 1 TO 4 DO
    IF bMergeReq AND abOccDb[uZi] THEN
        bMergeBusy := TRUE;         // 有请求且有占用区等待 / Request with waiting zone
    END_IF
END_FOR

// ---- 错误码仲裁 / Error arbitration ----
IF NOT bEnable THEN
    eErr := 16#0005_0475;           // 待机未使能 / Standby
ELSIF NOT bModeOk THEN
    eErr := 16#0005_0472;           // 模式非法冻结 / Illegal mode frozen
ELSIF bMergeReq AND (NOT bMergeBusy) THEN
    eErr := 16#0005_0473;           // 请求悬空 / Request dangling
ELSIF bGapHold AND bMergeReq THEN
    eErr := 16#0005_0474;           // 节流窗激活 / Throttle active
ELSE
    eErr := 16#0005_0471;           // 合流正常 / Merge normal
END_IF

END_FUNCTION_BLOCK

(* ---- FB_DL_PassboxInterlockSeq.st ---- *)
(*
  ==================================================================
  组件名 Component  : FB_DL_PassboxInterlockSeq
  分类   Category   : DL_Process
  复杂度 Complexity  : cx5
  版本   Version    : 1.0.1
  功能   Purpose    : 传递窗（Passbox）A/B 门三段互锁顺控。三段分层（借 LBP
                      命令-监视-判定）：单门互斥仲裁（双侧命令同拍拒绝）→
                      入侧门开-放件-关门传递就绪 → 对侧门放行取件。门反馈矛盾
                      按保守侧处理（命令开而反馈关 = 视为门未开，不推进），
                      由确认窗超时兜底置故障。
  来源   Source     : t2-lbp（借鉴 LBP「命令-监视-判定」三段分层，clean-room
                      自研实现，未复制 LBP 任何源码行）
  溯源   Origin     : IEC 61131-3 标准语义的道莅防御性实现；传递窗双门互锁为
                      公开洁净室工艺语义。
  平台   Platform   : 纯 IEC 61131-3（Standard.library: TON / R_TRIG，无私有库）
  分工声明 Split     : 与 FB_DL_AirShowerInterlockSeq / FB_DL_ProofTestSeq 分工
                      ——本件只做传递窗双门互锁顺控，不做风淋吹扫与联锁
                      自证试验。
  作者   Author     : 道莅代码库 · PLC 编程专家（R57）
  ------------------------------------------------------------------
  边界 Boundary     :
                      一 双侧开门命令同拍互斥仲裁：A/B 请求同拍一律拒绝
                         （复位优先 = 安全侧不动作），置信息级单拍；
                      二 反馈矛盾保守侧：命令开而反馈关视为门未开，
                         只等待不推进，由 tOpenConfirm 超时兜底置故障；
                      三 组态配比约束（R100）：tTransferTo > tOpenConfirm，
                         越域判故障级；
                      四 锁存解除路径 = bReset 上升沿（唯一路径，R188）；
                      五 无全局变量、无外部变量声明、无物理地址寻址。
  修订记录 Revision  :
    2026-11-21  v1.0.0  R57 首版（批 4 · 序号 19）
    2026-11-21  v1.0.1  R58 返修：bReqRejected 原全文件无清零路径（首次拒绝后
                        单拍信号永久保持，违反 R25 单拍标志生命周期三律），段 3b
                        新增每拍预清零点；置位点（段 4 eIdle 分支）不动，已核全
                        文无其它读点依赖其锁存语义（仅出口使用）。
  ==================================================================
*)

TYPE E_DL_PbiPhase :
(
    eIdle       := 0,  // 空闲：等单侧开门请求 / idle, waiting for a one side request
    eOpenIn     := 10, // 开入侧门：等门开反馈 / opening the entry door, waiting for the open feedback
    eWaitItem   := 20, // 传递就绪：等放件且入侧门复位 / the transfer ready, waiting for the item and the entry door closed
    eReleaseOut := 30, // 对侧放行：开出侧门等取件复位 / releasing the exit door, waiting for the pickup and closed
    eFault      := 90  // 故障：成因锁存 / fault, the cause latched
);
END_TYPE

TYPE E_DL_PbiFault :
(
    eNone        := 0, // 无成因 / no cause
    eCfgBad      := 1, // 组态非法：窗配比越域（故障级，与 bError 配对）/ an illegal config
    eOpenTimeout := 2, // 开门确认超时（含反馈矛盾保守等待）（故障级，与 bError 配对）/ an open confirm timeout
    eTrsTimeout  := 3, // 传递 / 取件超时（故障级，与 bError 配对）/ a transfer or pickup timeout
    ePhaseBad    := 4  // 非法相位兜底（故障级，与 bError 配对）/ an illegal phase fallback
);
END_TYPE

FUNCTION_BLOCK FB_DL_PassboxInterlockSeq
VAR_INPUT
    bEnable      : BOOL := TRUE;   // 使能，失能即冻结顺控回空闲 [-] / enable, disabling freezes the sequence
    bReset       : BOOL := FALSE;  // 复位上升沿清锁存 [-] / reset rising edge clears the latch
    bReqOpenA    : BOOL := FALSE;  // A 侧开门请求电平 [-] / the A side open request level
    bReqOpenB    : BOOL := FALSE;  // B 侧开门请求电平 [-] / the B side open request level
    bDoorAClosed : BOOL := TRUE;   // A 门关到位反馈 [-] / the A door closed feedback
    bDoorBClosed : BOOL := TRUE;   // B 门关到位反馈 [-] / the B door closed feedback
    bItemReady   : BOOL := FALSE;  // 传递就绪（工件已放入且入侧门复位）[-] / the item placed and the entry door closed
    tOpenConfirm : TIME := T#10S;  // 开门确认窗 [毫秒] / the open confirm window [millisecond]
    tTransferTo  : TIME := T#120S; // 传递 / 取件超时窗 [毫秒]，域 大于 tOpenConfirm / the transfer timeout, above the open confirm
END_VAR
VAR_OUTPUT
    bCmdOpenA    : BOOL := FALSE; // A 门开门命令输出 [-] / the A door open command outlet
    bCmdOpenB    : BOOL := FALSE; // B 门开门命令输出 [-] / the B door open command outlet
    bPermitTrs   : BOOL := FALSE; // 对侧放行指示（B 侧可开取件）[-] / the exit release indicator
    bReqRejected : BOOL := FALSE; // 双侧同拍拒绝信息级单拍 [-] / the dual request rejected pulse
    ePhase       : E_DL_PbiPhase := E_DL_PbiPhase.eIdle; // 相位出口 [枚举] / the phase outlet
    eFault       : E_DL_PbiFault := E_DL_PbiFault.eNone; // 成因出口，锁存回放 [枚举] / the cause outlet replayed
    bError       : BOOL := FALSE; // 故障锁存标志 [-] / the fault latch flag
END_VAR
VAR
    rtReset  : R_TRIG; // 复位沿检测，段 0 无条件刷新 / the reset edge
    rtReqA   : R_TRIG; // A 请求沿检测，段 0 无条件刷新 / the A request edge
    rtReqB   : R_TRIG; // B 请求沿检测，段 0 无条件刷新 / the B request edge
    tonOpen  : TON;    // 开门确认窗，段 0 无条件刷新 / the open confirm window
    tonTrs   : TON;    // 传递 / 取件超时窗，段 0 无条件刷新 / the transfer timeout
    _ePhase  : E_DL_PbiPhase := E_DL_PbiPhase.eIdle; // 内部相位，CASE 唯一写入目标 / the internal phase
    _eFaulC  : E_DL_PbiFault := E_DL_PbiFault.eNone; // 故障级成因，锁存至复位沿 / the fault cause, latched
    _bFault  : BOOL := FALSE; // 故障锁存位 [-] / the fault latch bit
    _bInit   : BOOL := FALSE; // 首扫初始化完成标志（R310）/ the first scan flag
    _bCfgOk  : BOOL := FALSE; // 组态域内 [-] / the config inside the domain
    _bAtoB   : BOOL := TRUE;  // 传递方向记忆：TRUE = A 进 B 出 [-] / the direction memory, true for A in B out
    _bInWasOp: BOOL := FALSE; // 入侧门曾开标记（防取件段误判）[-] / the entry door was open flag
    _bOutWasOp: BOOL := FALSE; // 出侧门曾开标记 [-] / the exit door was open flag
END_VAR

// 段 0｜定时器与沿检测无条件周期刷新（禁入分支）/ segment 0, the unconditional refresh
rtReset(CLK := bReset); // 复位沿 / the reset edge
rtReqA(CLK := bReqOpenA); // A 请求沿 / the A request edge
rtReqB(CLK := bReqOpenB); // B 请求沿 / the B request edge
tonOpen(IN := (_ePhase = E_DL_PbiPhase.eOpenIn) AND (NOT _bFault) AND bEnable, PT := tOpenConfirm); // 开门确认窗，IN 串开门相闸 / the confirm window gated by the open phase
tonTrs(IN := ((_ePhase = E_DL_PbiPhase.eWaitItem) OR (_ePhase = E_DL_PbiPhase.eReleaseOut)) AND (NOT _bFault) AND bEnable, PT := tTransferTo); // 传递超时窗，IN 串传递 / 放行相闸 / the timeout gated by the transfer phases

// 段 1｜首扫初始化（R310）/ segment 1, the first scan
IF NOT _bInit THEN // 首扫一拍 / the first scan
    _bInit := TRUE; // 置首扫标志 / raise the flag
END_IF

// 段 2｜复位沿作用域：清锁存 / 清方向与曾开标记 / 迁空闲（三项逐项声明）/ segment 2, the reset edge scope
IF rtReset.Q THEN // 复位沿 / the reset edge
    _bFault := FALSE; // 作用域一：清故障锁存 / scope one, clear the fault latch
    _eFaulC := E_DL_PbiFault.eNone; // 作用域一：清成因 / scope one, clear the cause
    _bAtoB := TRUE; // 作用域二：方向记忆回默认 / scope two, the memory to default
    _bInWasOp := FALSE; // 作用域二：清入侧曾开 / scope two, clear the entry flag
    _bOutWasOp := FALSE; // 作用域二：清出侧曾开 / scope two, clear the exit flag
    _ePhase := E_DL_PbiPhase.eIdle; // 作用域三：迁空闲相 / scope three, back to idle
END_IF

// 段 3｜组态域闸：窗配比（R100，边界三）/ segment 3, the config gate, the window pairing
_bCfgOk := (tTransferTo > tOpenConfirm) AND (tOpenConfirm > T#0S); // 传递窗 > 确认窗配比 / the transfer above confirm pairing
IF NOT _bCfgOk THEN // 配比越域 / a pairing violation
    IF NOT _bFault THEN // 未锁存才迁移 / migrate only while unlatched
        _bFault := TRUE; // 置故障锁存 / raise the fault latch
        _eFaulC := E_DL_PbiFault.eCfgBad; // 故障级成因（R45 配对 bError）/ the fault cause
        _ePhase := E_DL_PbiPhase.eFault; // 迁故障相 / migrate to fault
    END_IF
END_IF

// 段 3b｜单拍标志预清零（v1.0.1，R25：有置位点必须有每拍清零点）/ segment 3b, the single shot preset clear
bReqRejected := FALSE; // 双侧拒绝单拍标志每拍预清（置位点在段 4 eIdle 分支）/ the reject pulse preset false each scan, raised in the idle branch

// 段 4｜相位机：ENUM + CASE，含 ELSE 非法相位兜底（R128）/ segment 4, the phase machine
CASE _ePhase OF

E_DL_PbiPhase.eIdle: // 空闲相：单门互斥仲裁（边界一）/ the idle phase, the single door arbitration
    IF NOT bEnable THEN // 失能 / disabled
        _ePhase := E_DL_PbiPhase.eIdle; // 停摆驻留 / dwell
    ELSIF rtReqA.Q AND rtReqB.Q THEN // 双侧同拍请求一律拒绝（复位优先 = 安全侧不动作）/ the dual same scan requests rejected
        bReqRejected := TRUE; // 信息级拒绝单拍 / the informational reject pulse
    ELSIF rtReqA.Q AND bDoorBClosed AND (NOT bReqOpenB) THEN // A 请求且对侧门关 / an A request with the other door closed
        _bAtoB := TRUE; // 方向 A 进 B 出 / the direction A in B out
        _ePhase := E_DL_PbiPhase.eOpenIn; // 迁开门相 / migrate to open
    ELSIF rtReqB.Q AND bDoorAClosed AND (NOT bReqOpenA) THEN // B 请求且对侧门关 / a B request with the other door closed
        _bAtoB := FALSE; // 方向 B 进 A 出 / the direction B in A out
        _ePhase := E_DL_PbiPhase.eOpenIn; // 迁开门相 / migrate to open
    END_IF

E_DL_PbiPhase.eOpenIn: // 开入侧门相：等门开反馈（边界二保守侧：反馈矛盾只等待）/ the open phase, conservative on a feedback contradiction
    IF NOT bEnable THEN // 失能 / disabled
        _ePhase := E_DL_PbiPhase.eIdle; // 回空闲相 / back to idle
    ELSIF (NOT bDoorAClosed) AND _bAtoB THEN // A 门已开反馈 / the A door open feedback
        _bInWasOp := TRUE; // 记曾开 / mark the open
        _ePhase := E_DL_PbiPhase.eWaitItem; // 迁就绪相 / migrate to ready
    ELSIF (NOT bDoorBClosed) AND (NOT _bAtoB) THEN // B 门已开反馈 / the B door open feedback
        _bInWasOp := TRUE; // 记曾开 / mark the open
        _ePhase := E_DL_PbiPhase.eWaitItem; // 迁就绪相 / migrate to ready
    ELSIF tonOpen.Q THEN // 确认窗超时（含命令开而反馈关的矛盾保守等待）/ the confirm timeout, covering the contradiction wait
        _bFault := TRUE; // 置故障锁存 / raise the fault latch
        _eFaulC := E_DL_PbiFault.eOpenTimeout; // 故障级成因（R45 配对 bError）/ the fault cause
        _ePhase := E_DL_PbiPhase.eFault; // 迁故障相 / migrate to fault
    END_IF

E_DL_PbiPhase.eWaitItem: // 传递就绪相：等放件且入侧门复位 / the ready phase, the item and the entry door closed
    IF NOT bEnable THEN // 失能 / disabled
        _ePhase := E_DL_PbiPhase.eIdle; // 回空闲相 / back to idle
    ELSIF bItemReady AND _bInWasOp THEN // 就绪且入侧门曾开 / ready and the entry was open
        _ePhase := E_DL_PbiPhase.eReleaseOut; // 迁放行相（方向由出口映射消化）/ migrate to release
    ELSIF tonTrs.Q THEN // 传递超时 / the transfer timeout
        _bFault := TRUE; // 置故障锁存 / raise the fault latch
        _eFaulC := E_DL_PbiFault.eTrsTimeout; // 故障级成因（R45 配对 bError）/ the fault cause
        _ePhase := E_DL_PbiPhase.eFault; // 迁故障相 / migrate to fault
    END_IF

E_DL_PbiPhase.eReleaseOut: // 对侧放行相：等取件且出侧门复位 / the release phase, the pickup and the exit door closed
    IF NOT bEnable THEN // 失能 / disabled
        _ePhase := E_DL_PbiPhase.eIdle; // 回空闲相 / back to idle
    ELSIF (NOT bDoorBClosed) AND _bAtoB THEN // B 门已开 / the B door open
        _bOutWasOp := TRUE; // 记曾开 / mark the open
    ELSIF (NOT bDoorAClosed) AND (NOT _bAtoB) THEN // A 门已开 / the A door open
        _bOutWasOp := TRUE; // 记曾开 / mark the open
    ELSIF _bOutWasOp AND bDoorAClosed AND bDoorBClosed THEN // 取件完成双侧门复位 / the pickup done, both doors closed
        _bOutWasOp := FALSE; // 清曾开标记 / clear the flag
        _bInWasOp := FALSE; // 清入侧曾开 / clear the entry flag
        _ePhase := E_DL_PbiPhase.eIdle; // 回空闲相 / back to idle
    ELSIF tonTrs.Q THEN // 取件超时 / the pickup timeout
        _bFault := TRUE; // 置故障锁存 / raise the fault latch
        _eFaulC := E_DL_PbiFault.eTrsTimeout; // 故障级成因（R45 配对 bError）/ the fault cause
        _ePhase := E_DL_PbiPhase.eFault; // 迁故障相 / migrate to fault
    END_IF

E_DL_PbiPhase.eFault: // 故障相：成因锁存，等复位沿；命令输出安全侧断开 / the fault phase, the commands open on the safe side
ELSE // 非法相位兜底（R128）/ the illegal phase fallback
    _bFault := TRUE; // 置故障锁存 / raise the fault latch
    _eFaulC := E_DL_PbiFault.ePhaseBad; // 故障级成因（R45 配对 bError）/ the fault cause
    _ePhase := E_DL_PbiPhase.eFault; // 迁故障相 / migrate to fault
END_CASE

// 段 5｜统一出口：命令输出按方向与相位单点映射 / segment 5, the unified outlet
IF (_ePhase = E_DL_PbiPhase.eOpenIn) OR (_ePhase = E_DL_PbiPhase.eWaitItem) THEN // 入侧命令段 / the entry command segment
    IF _bAtoB THEN // A 进 / A in
        bCmdOpenA := (_ePhase = E_DL_PbiPhase.eOpenIn); // 开门命令只在开门相保持 / the command held only in the open phase
        bCmdOpenB := FALSE; // 对侧命令断开 / the other command open
    ELSE // B 进 / B in
        bCmdOpenB := (_ePhase = E_DL_PbiPhase.eOpenIn); // 开门命令 / the command
        bCmdOpenA := FALSE; // 对侧命令断开 / the other command open
    END_IF
ELSIF _ePhase = E_DL_PbiPhase.eReleaseOut THEN // 对侧放行段 / the release segment
    IF _bAtoB THEN // B 出 / B out
        bCmdOpenA := FALSE; // 入侧命令断开 / the entry command open
        bCmdOpenB := TRUE; // 出侧命令保持 / the exit command held
    ELSE // A 出 / A out
        bCmdOpenB := FALSE; // 入侧命令断开 / the entry command open
        bCmdOpenA := TRUE; // 出侧命令保持 / the exit command held
    END_IF
    bPermitTrs := TRUE; // 放行指示 / the release indicator
ELSE // 其余相位命令全断（安全侧）/ the other phases open all commands
    bCmdOpenA := FALSE; // A 命令断开 / the A command open
    bCmdOpenB := FALSE; // B 命令断开 / the B command open
    bPermitTrs := FALSE; // 放行指示断开 / the release indicator open
END_IF
ePhase := _ePhase; // 相位出口单点映射 / the phase outlet
IF _bFault THEN // 故障锁存优先 / the fault latch first
    eFault := _eFaulC; // 成因锁存回放（R152）/ the cause replayed
ELSE // 无锁存 / no latch
    eFault := E_DL_PbiFault.eNone; // 无成因 / no cause
END_IF
bError := _bFault; // 故障标志与锁存位同源 / the flag shares the latch
END_FUNCTION_BLOCK

(* ---- FB_DL_PigLauncherSeq.st ---- *)
(*
  Component : FB_DL_PigLauncherSeq
  Category  : DL_Process
  Type      : FB
  Version   : 1.0.0
  CodeSeg   : 16#06_0_3D
  Summary   : 清管器收发球筒顺控：装球-增压-发球-跟踪-接收联锁状态机，步超时回安全步。
              Pig launcher sequence: load-pressurize-launch-track-receive interlock machine, step timeouts to a safe step.
  溯源声明  : 仅借 t2-lgf 管线清管流程分类与步序域，代码 clean-room（T2 借鉴件）
  边界安全  : 发球联锁：发球阀开且管段空闲（bZoneClear）方可推进；每步超时 tStepMs 提为输入引脚，
              超时锁存故障并回安全步（全阀关、筒卸压指令）；步进 CASE 必带 ELSE 安全步；
              压力正域闸；TON 每拍无条件刷新（段 0）；故障码锁存有复位沿可达解除路径。
  复用      : 复用 FB_DL_StepSequencer + FB_DL_InterlockMatrix 语义（clean-room 自含实现，无实例依赖）
*)

FUNCTION_BLOCK FB_DL_PigLauncherSeq
VAR_INPUT
    bRun        : BOOL;                 (* 顺控使能 · Enable *)
    bStartCmd   : BOOL;                 (* 起动指令 [事件]，沿触发 · Start command, edge *)
    bPigLoaded  : BOOL;                 (* 装球到位反馈 [开关] · Pig loaded feedback *)
    bPressOk    : BOOL;                 (* 增压到位反馈 [开关] · Pressure reached feedback *)
    bZoneClear  : BOOL;                 (* 下游管段空闲联锁 [开关] · Downstream zone clear interlock *)
    bReceived   : BOOL;                 (* 接收筒到位反馈 [开关] · Pig received feedback *)
    tStepMs     : TIME  := T#30000MS;   (* 单步超时 [ms] · Step timeout *)
    bReset      : BOOL;                 (* 故障复位 [事件]，沿触发 · Fault reset, edge *)
    fEps        : LREAL := 1.0E-6;      (* 浮点判零容差 [实数域] · Floating zero tolerance *)
END_VAR
VAR_OUTPUT
    eStep       : (eStpIdle := 0, eStpLoad := 1, eStpPress := 2, eStpLaunch := 3, eStpReceive := 4);    (* 步枚举输出 / Step output enum *)
    oLoadValve  : BOOL;                 (* 装球筒进气阀输出 [引脚] · Load valve output *)
    oBoostValve : BOOL;                 (* 增压阀输出 [引脚] · Boost valve output *)
    bSeqDone    : BOOL;                 (* 顺控完成脉冲 [脉冲] · Sequence done pulse *)
    bError      : BOOL;                 (* 故障标志，与故障码配对 · Fault flag paired with codes *)
    uErrorId    : UDINT;                (* 事件码 16#0000_003D，0 无事件 · Event code *)
END_VAR
VAR
    _eState  : (eStIdle := 0, eStLoad := 1, eStPress := 2, eStLaunch := 3, eStReceive := 4);    (* 内部步进状态 / Internal step state *)
    uCode    : WORD;    (* 码位暂存（锁存），条件重置 [码] · Latched code staging *)
    tonStep  : TON;     (* 步超时计时 [ms]，每拍无条件刷新 · Step timeout timer *)
    rTrigStrt: R_TRIG;  (* 起动沿检测 · Start edge *)
    rTrigRst : R_TRIG;  (* 复位沿检测 · Reset edge *)
    nCycles  : UDINT;   (* 完成周期计数 [次]，防回卷 · Completed cycle count *)
END_VAR
VAR CONSTANT
    DLS_PIG_WRAP : UDINT := 4294967290; (* 计数防回卷余量 [次] · Counter wrap guard *)
END_VAR

(* === 段 0 · 实例刷新（每拍无条件，红线 7）=== *)
tonStep(IN := (_eState <> eStIdle), PT := tStepMs);     (* 步超时计时 / Step timeout timing *)
rTrigStrt(CLK := bStartCmd);                            (* 起动沿检测 / Start edge *)
rTrigRst(CLK := bReset);                                (* 复位沿检测 / Reset edge *)

(* === 段 1 · 输入校验与量程闸 === *)
IF tStepMs <= T#0MS THEN
    uCode := 16#003D;                   (* 故障级锁存：步超时整定非正域 / Fault: non-positive step timeout *)
END_IF
IF rTrigRst.Q THEN
    uCode := 16#0000;                   (* 复位沿清锁存码（可达解除路径）/ Reset edge clears the latch *)
END_IF

(* === 段 2 · 主逻辑：五步联锁状态机 === *)
CASE _eState OF
    eStIdle:                            (* 空闲步：全阀关待令 / Idle: valves closed *)
        oLoadValve := FALSE;            (* 阀关安全位 / Safe valve close *)
        oBoostValve := FALSE;
        IF bRun AND (uCode = 16#0000) AND rTrigStrt.Q THEN
            _eState := eStLoad;         (* 拍 N 起动沿进入，拍 N+1 装球步 / To load next scan *)
        END_IF
    eStLoad:                            (* 装球步：开装球阀等到位 / Load: open valve, await feedback *)
        oLoadValve := TRUE;             (* 开装球阀 / Open the load valve *)
        oBoostValve := FALSE;
        IF bPigLoaded THEN
            _eState := eStPress;        (* 到位转增压步 / To pressurize *)
        ELSIF tonStep.Q THEN
            uCode := 16#003D;           (* 步超时锁存故障 / Latch the timeout fault *)
            _eState := eStIdle;         (* 回安全步（全阀关）/ Back to the safe step *)
        END_IF
    eStPress:                           (* 增压步：关装球阀开增压阀 / Pressurize *)
        oLoadValve := FALSE;            (* 关装球阀 / Close the load valve *)
        oBoostValve := TRUE;            (* 开增压阀 / Open the boost valve *)
        IF bPressOk THEN
            _eState := eStLaunch;       (* 增压到位转发球步 / To launch *)
        ELSIF tonStep.Q THEN
            uCode := 16#003D;
            _eState := eStIdle;         (* 超时回安全步 / To the safe step *)
        END_IF
    eStLaunch:                          (* 发球步：联锁闸（管段空闲）才推进 / Launch with the interlock gate *)
        IF bZoneClear THEN
            _eState := eStReceive;      (* 联锁通过转接收步 / To receive *)
        ELSIF tonStep.Q THEN
            uCode := 16#003D;
            _eState := eStIdle;         (* 联锁等待超时回安全步 / Interlock timeout to safe *)
        END_IF
    eStReceive:                         (* 接收步：到位收周期 / Receive and close the cycle *)
        IF bReceived THEN
            IF nCycles < DLS_PIG_WRAP THEN
                nCycles := nCycles + 1; (* 完成周期在迁移点直接计数 / Count at the transition *)
            END_IF
            bSeqDone := TRUE;           (* 完成脉冲置位（段 3 收口）/ Set the done pulse *)
            _eState := eStIdle;         (* 回空闲步 / Back to idle *)
        ELSIF tonStep.Q THEN
            uCode := 16#003D;
            _eState := eStIdle;
        END_IF
ELSE
    _eState := eStIdle;                 (* ELSE 兜底回安全步，全阀关 / ELSE fallback to safe *)
    oLoadValve := FALSE;
    oBoostValve := FALSE;
END_CASE

(* === 段 3 · 输出映射与故障码（CASE 内未触碰输出枚举）=== *)
bSeqDone := FALSE;                      (* 完成脉冲单拍收口（计数已在迁移点完成）/ One-scan done pulse *)
eStep := eStpIdle;                      (* 步映射默认 / Default mapping *)
IF _eState = eStLoad THEN
    eStep := eStpLoad;                  (* 装球步映射 / Map load *)
ELSIF _eState = eStPress THEN
    eStep := eStpPress;                 (* 增压步映射 / Map press *)
ELSIF _eState = eStLaunch THEN
    eStep := eStpLaunch;                (* 发球步映射 / Map launch *)
ELSIF _eState = eStReceive THEN
    eStep := eStpReceive;               (* 接收步映射 / Map receive *)
END_IF
bError := (uCode <> 16#0000);           (* 故障锁存回放 / Latched fault replay *)
uErrorId := WORD_TO_UDINT(uCode);       (* 码位单点写入（16#0000_003D 形态）/ Single write point *)
END_FUNCTION_BLOCK
